IF _n > 0 THEN
    _n          := _n - 1;
    stsVerified := FALSE;
    IF _n = 0 THEN
        _state := E_CamTeach_State.eIdle;
    ELSE
        _state := eTeaching;
    END_IF
END_IF
cmdDeleteLast := TRUE;
END_METHOD

// Spot-edit one existing point (offline, before convert/download). Clears verified.
// Faults on an out-of-range index. Rejected QUIETLY while busy/errored.
METHOD PUBLIC cmdEditPoint : BOOL
VAR_INPUT
    idx     : INT;     // 1..stsNumPoints
    rMaster : LREAL;   // [master unit] new master value
    rSlave  : LREAL;   // [slave unit]  new slave value
END_VAR
cmdEditPoint := FALSE;
IF isBusy() OR stsError THEN
    RETURN;
END_IF

IF idx < 1 OR idx > _n THEN
    setError('Edit point: index out of range');
    RETURN;
END_IF

_points[idx].rMaster := rMaster;
_points[idx].rSlave  := rSlave;
stsVerified  := FALSE;
_state       := eTeaching;
cmdEditPoint := TRUE;
END_METHOD

// Empty the working set (returns toward E_CamTeach_State.eIdle). Clears verified. Rejected QUIETLY while busy/errored.
METHOD PUBLIC cmdClear : BOOL
cmdClear := FALSE;
IF isBusy() OR stsError THEN
    RETURN;
END_IF

_n          := 0;
stsVerified := FALSE;
_state      := E_CamTeach_State.eIdle;
cmdClear    := TRUE;
END_METHOD

// Persist the raw points -> file (async, via fb_CamTeachFile). The directory is cfgFileDir;
// the caller passes just a bare file name. Metadata (slaveName/created/periodic/interp/masterUnit)
// is taken from the cfg backing except 'created', which the HMI stamps (wall clock not in-scan).
// Rejected QUIETLY while busy/errored or with nothing to save.
METHOD PUBLIC cmdSave : BOOL
VAR_INPUT
    fileName : STRING;   // bare file name, e.g. '<pattern>_<slaveName>.csv'
END_VAR
VAR
    sInterp : STRING;
END_VAR
cmdSave := FALSE;
IF isBusy() OR stsError THEN
    RETURN;
END_IF

IF _n < 1 THEN
    setError('Save: nothing to save');
    RETURN;
END_IF

// string form of the interpolation strategy for the CSV '#' header
sInterp := SEL(_interp = E_CamTeach_Interp.eCubicC1, 'linear', 'cubicC1');

IF _file.cmdSave(
        dir        := _fileDir,
        fileName   := fileName,
        numPoints  := _n,
        slaveName  := _slaveName,
        created    := HMI.Config.created,
        periodic   := _periodic,
        interp     := sInterp,
        masterUnit := _masterUnit) THEN
    _fileName    := fileName;
    _returnState := _state;         // resting state to return to once the write completes
    _state       := eSaving;
    cmdSave      := TRUE;
END_IF
END_METHOD

// File -> raw points (async, via fb_CamTeachFile). On completion _n is taken from
// _file.stsNumPointsLoaded and validated (>= 2) in the eLoading branch of the body.
// Loading invalidates any verified table. Rejected QUIETLY while busy/errored.
METHOD PUBLIC cmdLoad : BOOL
VAR_INPUT
    fileName : STRING;   // bare file name to load (directory is cfgFileDir)
END_VAR
cmdLoad := FALSE;
IF isBusy() OR stsError THEN
    RETURN;
END_IF

IF _file.cmdLoad(dir := _fileDir, fileName := fileName) THEN
    _fileName := fileName;
    _state    := eLoading;
    cmdLoad   := TRUE;
END_IF
END_METHOD

// SYNCHRONOUS: post-process the raw points then build the NC motion function _mfPoints[].
// Pure and bounded by MAX_CAM_POINTS (no I/O), so it completes in one scan -> eConverted.
// Post-processing is IN PLACE (design doc "compact the array"): it zeroes the master offset,
// deletes non-monotonic points, and optionally smooths the master column, updating _n. Save
// the raw points BEFORE converting if the untouched values are needed. A (re)convert also
// invalidates any prior download (stsVerified := FALSE). Rejected QUIETLY while busy/errored.
METHOD PUBLIC cmdConvert : BOOL
VAR
    base : LREAL;   // master offset removed in step 1
    i    : INT;     // point loop index
    j    : INT;     // compaction write cursor
    w2   : INT;     // smoothing half-window
    lo   : INT;     // smoothing window low bound
    hi   : INT;     // smoothing window high bound
    k    : INT;     // smoothing inner index
    sum  : LREAL;   // smoothing accumulator
END_VAR
cmdConvert := FALSE;
IF isBusy() OR stsError THEN
    RETURN;
END_IF

IF _n < 2 THEN
    setError('Convert: need at least 2 taught points');
    RETURN;
END_IF

// A (re)convert invalidates any previously downloaded/verified table.
stsVerified := FALSE;

// ── Post-processing 1: zero the master offset (table starts at master = 0) ──
base := _points[1].rMaster;
FOR i := 1 TO _n DO
    _points[i].rMaster := _points[i].rMaster - base;
END_FOR

// ── Post-processing 2: enforce strict-monotonic master (compact the array in place) ──
// Keep point 1; keep each later point only if its master exceeds the last kept point's.
j := 1;
FOR i := 2 TO _n DO
    IF _points[i].rMaster > _points[j].rMaster THEN
        j := j + 1;
        _points[j] := _points[i];
    END_IF
END_FOR
_n := j;
IF _n < 2 THEN
    setError('Convert: too few monotonic points');
    RETURN;
END_IF

// ── Post-processing 3: optional moving-average smoothing of the MASTER column ──
// Odd window (>= 3); the window shrinks at the endpoints. _mfPoints[].MasterPos is used as
// scratch so each average is taken from the ORIGINAL masters (an in-place average would feed
// already-smoothed neighbours into later points). 0/1/2 disable smoothing.
IF _smoothWindow >= 3 THEN
    w2 := (_smoothWindow - 1) / 2;
    FOR i := 1 TO _n DO
        lo := i - w2;  IF lo < 1  THEN lo := 1;  END_IF
        hi := i + w2;  IF hi > _n THEN hi := _n; END_IF
        sum := 0.0;
        FOR k := lo TO hi DO
            sum := sum + _points[k].rMaster;
        END_FOR
        _mfPoints[i].MasterPos := sum / INT_TO_LREAL(hi - lo + 1);   // scratch (overwritten below)
    END_FOR
    FOR i := 1 TO _n DO
        _points[i].rMaster := _mfPoints[i].MasterPos;
    END_FOR
END_IF

// ── Build the NC motion function (C1-smooth cubic from position-only teaching) ──
// Field names and enums checked against TF5050 manual 1.9.2 (section 9.7-9.10), 2026-10-18.
// PointType MUST be set: its default 0 is MOTIONPOINTTYPE_IGNORE, and a table of ignored points is
// rejected (NC 0x4A23 'Motion Function has too few points'). Segments are POLYNOM3_VV (velo <-> velo:
// a cubic through each point's position AND slope) - plain POLYNOM3 is rest <-> rest, i.e. the slave
// would stop at every taught point whatever SlaveVelo says.
FOR i := 1 TO _n DO
    _mfPoints[i].PointIndex        := INT_TO_UDINT(i);       // 1, 2, 3 ... (> 0, consecutive, no gaps)
    _mfPoints[i].PointType         := MOTIONPOINTTYPE_MOTION;
    _mfPoints[i].RelIndexNextPoint := 1;
    _mfPoints[i].MasterPos         := _points[i].rMaster;
    _mfPoints[i].SlavePos          := _points[i].rSlave;
    _mfPoints[i].SlaveVelo         := slaveSlope(i);         // dSlave/dMaster at this point
    _mfPoints[i].SlaveAcc          := 0.0;
    _mfPoints[i].SlaveJerk         := 0.0;
    IF i = _n THEN
        _mfPoints[i].FunctionType      := MOTIONFUNCTYPE_NOTDEF; // last point: no segment after it
        _mfPoints[i].RelIndexNextPoint := 0;                     // ... and no next point (1 -> index _n+1, NC 0x4A13?)
    ELSE
        _mfPoints[i].FunctionType := MOTIONFUNCTYPE_POLYNOM3_VV; // segment to the next point
    END_IF
END_FOR

_state     := eConverted;
cmdConvert := TRUE;
END_METHOD

// Start the async download -> verify state machine (MC_CamTableSelect creates the table, then per-point
// MC_ReadMotionFunctionPoint read-back). On success -> eVerified + stsVerified := TRUE. Requires
// eConverted and a bound cfgTableId. Rejected QUIETLY while busy/errored.
METHOD PUBLIC cmdDownload : BOOL
cmdDownload := FALSE;
IF isBusy() OR stsError THEN
    RETURN;
END_IF

IF _state <> eConverted THEN
    setError('Download: convert first (must be in eConverted)');
    RETURN;
END_IF

IF _tableId = 0 THEN
    setError('Download: no NC cam table id configured');
    RETURN;
END_IF

IF _n < 2 THEN
    setError('Download: nothing to download');
    RETURN;
END_IF

stsVerified := FALSE;               // clears any prior verify until this download re-verifies
_dlStep     := 0;
_state      := eDownloading;
cmdDownload := TRUE;
END_METHOD

// Live single-point slave edit while the table is in use. Updates _points[idx].rSlave, rebuilds
// the affected motion-function points (the edited point's SlavePos + the slopes of it and its
// immediate neighbours), then kicks the async sequence: set the online-change mode (apply at a
// defined master position, NOT immediately) and write the affected points via
// MC_WriteMotionFunctionPoint. The file is re-saved so it stays truthful. A live edit clears
// stsVerified (a full re-convert + re-download is required before coupling is allowed again).
// Rejected QUIETLY while busy/errored, on a bad index, or with no bound table.
METHOD PUBLIC cmdEditOnline : BOOL
VAR_INPUT
    idx    : INT;     // 1..stsNumPoints target point index
    rSlave : LREAL;   // [slave unit] new slave value for the live edit
END_VAR
VAR
    k  : INT;
    lo : INT;
    hi : INT;
END_VAR
cmdEditOnline := FALSE;
IF isBusy() OR stsError THEN
    RETURN;
END_IF

IF _n < 2 THEN
    setError('Online edit: table too small');
    RETURN;
END_IF

IF idx < 1 OR idx > _n THEN
    setError('Online edit: index out of range');
    RETURN;
END_IF

IF _tableId = 0 THEN
    setError('Online edit: no NC cam table id configured');
    RETURN;
END_IF

// 1) update the working point and rebuild the affected motion-function points
//    (only the slave changed; recompute SlavePos of idx and the slopes of idx-1..idx+1).
_onlineIdx := idx;
_points[idx].rSlave := rSlave;

lo := idx - 1;  IF lo < 1  THEN lo := 1;  END_IF
hi := idx + 1;  IF hi > _n THEN hi := _n; END_IF
FOR k := lo TO hi DO
    _mfPoints[k].SlavePos  := _points[k].rSlave;    // VERIFY: MC_MotionFunctionPoint.SlavePos
    _mfPoints[k].SlaveVelo := slaveSlope(k);        // VERIFY: MC_MotionFunctionPoint.SlaveVelo
END_FOR

// 2) + 3) arm the async write sequence: change-mode first, then write points lo..hi.
_onlineWriteIdx := lo;
_onlineHi       := hi;
_onlineStep     := 10;
_onlineSaveReq  := TRUE;

// 4) a live edit invalidates the verified permission; report the updated-but-unverified state.
stsVerified := FALSE;
_state      := eConverted;

cmdEditOnline := TRUE;
END_METHOD

// Clear the FB's own error, reset the file sub-FB, and return to E_CamTeach_State.eIdle. Also aborts any in-flight
// download/verify/online sequence. stsVerified is cleared so a fresh convert + download + verify
// is required after a reset. Called from inpReset, ocmdReset, and directly.
METHOD PUBLIC cmdReset : BOOL
stsError     := FALSE;
stsErrorText := '';
_file.cmdReset();

_state          := E_CamTeach_State.eIdle;
_dlStep         := 0;
_verifyIdx      := 1;
_onlineStep     := 0;
_onlineWriteIdx := 1;
_onlineSaveReq  := FALSE;
stsVerified     := FALSE;
cmdReset        := TRUE;
END_METHOD

// Central-difference slave slope d(slave)/d(master) at point idx, used for the cubic SlaveVelo.
// Interior points use the central difference; the endpoints use one-sided differences. For a
// PERIODIC table the seam (point 1 == point _n phase) wraps so the slope is continuous across
// the period boundary. Assumes masters are strictly monotonic (post-processed); guards dM = 0.
METHOD PRIVATE slaveSlope : LREAL
VAR_INPUT
    idx : INT;     // 1.._n
END_VAR
VAR
    dM     : LREAL;
    dS     : LREAL;
    period : LREAL;
END_VAR
slaveSlope := 0.0;
IF _n < 2 OR idx < 1 OR idx > _n THEN
    RETURN;
END_IF

IF _periodic AND _n >= 3 AND (idx = 1 OR idx = _n) THEN
    // Seam wrap: _points[1] (master 0) and _points[_n] (master = period) are the SAME phase,
    // so idx=1 and idx=_n get the SAME (continuous) slope. period = the zeroed master span.
    period := _points[_n].rMaster - _points[1].rMaster;
    dS     := _points[2].rSlave - _points[_n - 1].rSlave;
    dM     := (_points[2].rMaster + period) - _points[_n - 1].rMaster;
ELSIF idx = 1 THEN
    // one-sided forward difference at the start
    dS := _points[2].rSlave  - _points[1].rSlave;
    dM := _points[2].rMaster - _points[1].rMaster;
ELSIF idx = _n THEN
    // one-sided backward difference at the end
    dS := _points[_n].rSlave  - _points[_n - 1].rSlave;
    dM := _points[_n].rMaster - _points[_n - 1].rMaster;
ELSE
    // interior central difference
    dS := _points[idx + 1].rSlave  - _points[idx - 1].rSlave;
    dM := _points[idx + 1].rMaster - _points[idx - 1].rMaster;
END_IF

IF dM <> 0.0 THEN
    slaveSlope := dS / dM;
END_IF
END_METHOD

// Latch the FB's own error (this FB does NOT extend abs_fb_Device - never setFault, which would
// gate MC_Power on a real axis). Moves to E_CamTeach_State.eError and aborts any in-flight download/verify/online
// sub-steps so the MC blocks de-assert next scan. Cleared only by cmdReset / inpReset.
METHOD PRIVATE setError : BOOL
VAR_INPUT
    text : STRING;
END_VAR
stsError     := TRUE;
stsErrorText := text;
_state       := E_CamTeach_State.eError;
_dlStep      := 0;
_onlineStep  := 0;
setError     := TRUE;
END_METHOD

// TRUE while any async operation is in progress (file save/load, download, verify, or online
// edit). Command methods use this to reject re-entrant requests without disturbing the running op.
METHOD PRIVATE isBusy : BOOL
isBusy := _file.stsBusy
    OR (_state = eSaving) OR (_state = eLoading)
    OR (_state = eDownloading) OR (_state = eVerifying)
    OR (_onlineStep <> 0);
END_METHOD

// Return the full HMI interface struct (the one an HMI binds).
METHOD PUBLIC getHMIdata : ST_CamTeach_HMI_Interface
getHMIdata := HMI;
END_METHOD

METHOD FB_Init : BOOL
VAR_INPUT
    bInitRetains    : BOOL;
    bInCopyCode     : BOOL;
    cfgTableId      : UDINT;              // NC motion-function table id bound to this instance
    cfgSlaveName    : STRING;             // name of the slave this table teaches (file header)
    cfgPeriodic     : BOOL;              // TRUE = periodic table (velocity wraps at the seam)
    cfgInterp       : E_CamTeach_Interp;  // interpolation strategy for cmdConvert
    cfgSmoothWindow : INT;               // moving-average window on master column (0 = off)
    cfgFileDir      : STRING;            // save/load directory ('' = keep default C:\_MachineConfig\CamTables)
    cfgMasterUnit   : STRING;            // CSV header master unit ('' = keep default 'mm')
END_VAR
_tableId   := cfgTableId;
_slaveName := cfgSlaveName;
_periodic  := cfgPeriodic;
_interp    := cfgInterp;
IF cfgSmoothWindow >= 0 THEN _smoothWindow := cfgSmoothWindow; END_IF
IF cfgFileDir    <> '' THEN _fileDir    := cfgFileDir;    END_IF
IF cfgMasterUnit <> '' THEN _masterUnit := cfgMasterUnit; END_IF
END_METHOD

// NC motion-function table id this instance downloads to (pre-created under Motion -> Tables).
PROPERTY PUBLIC cfgTableId : UDINT
GET
cfgTableId := _tableId;
END_GET
SET
_tableId := cfgTableId;
END_SET
END_PROPERTY

// Name of the slave this table teaches; written into the CSV '#' metadata header.
PROPERTY PUBLIC cfgSlaveName : STRING
GET
cfgSlaveName := _slaveName;
END_GET
SET
_slaveName := cfgSlaveName;
END_SET
END_PROPERTY

// TRUE = periodic table: the conversion wraps the central-difference slope at the seam so the
// slave velocity is continuous across the period boundary.
PROPERTY PUBLIC cfgPeriodic : BOOL
GET
cfgPeriodic := _periodic;
END_GET
SET
_periodic := cfgPeriodic;
END_SET
END_PROPERTY

// Interpolation strategy used by cmdConvert (eLinear / eCubicC1). eCubicC1 = POLYNOM3 +
// central-difference slope -> C1-smooth cubic from position-only teaching.
PROPERTY PUBLIC cfgInterp : E_CamTeach_Interp
GET
cfgInterp := _interp;
END_GET
SET
_interp := cfgInterp;
END_SET
END_PROPERTY

// Moving-average window applied to the master column in cmdConvert (odd, 3-5; 0 = off).
// A value < 0 is rejected; 1/2 act as off (the convert only smooths for windows >= 3).
PROPERTY PUBLIC cfgSmoothWindow : INT
GET
cfgSmoothWindow := _smoothWindow;
END_GET
SET
IF cfgSmoothWindow >= 0 THEN _smoothWindow := cfgSmoothWindow; END_IF
END_SET
END_PROPERTY

// Save/load directory (the caller passes only a bare file name). Default C:\_MachineConfig\CamTables.
PROPERTY PUBLIC cfgFileDir : STRING
GET
cfgFileDir := _fileDir;
END_GET
SET
IF cfgFileDir <> '' THEN _fileDir := cfgFileDir; END_IF
END_SET
END_PROPERTY

// Master unit label written into the CSV '#' header (e.g. 'mm' / 'deg'). Default 'mm'.
// Added beyond the design doc's cfg list because the file header needs a machine-specific
// master unit that fb_CamTeachFile.cmdSave requires (see the FB header note / report).
PROPERTY PUBLIC cfgMasterUnit : STRING
GET
cfgMasterUnit := _masterUnit;
END_GET
SET
IF cfgMasterUnit <> '' THEN _masterUnit := cfgMasterUnit; END_IF
END_SET
END_PROPERTY

END_FUNCTION_BLOCK

// ---- POUs/FBs/Camming/fb_CamTeachFile.TcPOU
// fb_CamTeachFile - isolated async CSV persistence for ONE cam-teach table.
//
// Standalone library primitive: does NOT extend abs_fb_Device. It carries its own
// error model (stsError / stsErrorId / stsErrorText) and is driven cyclically by
// fb_CamTeach, which passes its working point array in via VAR_IN_OUT every scan.
//
// The body mirrors the Tc2_System FB_File* async pattern (see fb_WriteDataToFile):
// FB_FileOpen -> FB_FilePuts / FB_FileGets -> FB_FileClose, sequenced by an nState
// CASE machine. Every step is non-blocking (one line per scan pass) and the error
// path (900..) ALWAYS closes the handle before halting.
//
// Operations are started ONLY from cmdSave / cmdLoad, and only when idle (nState = 0),
// so the body never self-triggers. The file is the source of truth; store RAW points.
//
// CSV format (raw values):
//   # slaveName=..  created=..  numPoints=..  periodic=0|1  interp=..  masterUnit=..
//   <master>, <slave>
//   ...
FUNCTION_BLOCK fb_CamTeachFile
VAR_IN_OUT
    // Shared working buffer owned by fb_CamTeach (passed in every scan).
    // Save reads points[1..numPoints]; Load overwrites points[1..stsNumPointsLoaded].
    points : ARRAY[1..MAX_CAM_POINTS] OF ST_CamTeach_Point;
END_VAR
VAR_OUTPUT
    stsBusy            : BOOL;    // an async save/load is in progress
    stsDone            : BOOL;    // last operation finished OK (latched until next op / cmdReset)
    stsError           : BOOL;    // last operation failed (latched until cmdReset)
    stsErrorId         : UDINT;   // Tc2 file-FB error id (nErrId) of the failing step, else 0
    stsErrorText       : STRING;  // human-readable failure description
    stsNumPointsLoaded : INT;     // number of points loaded by the last cmdLoad
END_VAR
VAR
    nState        : INT;          // 0 idle; 10.. save; 110.. load; 900.. error

    // Tc2_System line-oriented file blocks (async; one line per FB_FilePuts/FB_FileGets)
    fbFileOpen    : FB_FileOpen;
    fbFilePuts    : FB_FilePuts;
    fbFileGets    : FB_FileGets;
    fbFileClose   : FB_FileClose;
    hFile         : UINT := 0;    // open file handle (0 = closed)

    // Operation parameters captured by cmdSave / cmdLoad
    _dir          : STRING(255);
    _fileName     : STRING(255);
    _slaveName    : STRING;
    _created      : STRING;
    _interp       : STRING;
    _masterUnit   : STRING;
    _numPoints    : INT;          // points to save (from cmdSave)
    _periodic     : BOOL;

    // Working scratch
    sFullFilePath : STRING(255);  // dir + '\' + fileName
    sLine         : STRING(255);  // line buffer (built for puts / trimmed from gets)
    _i            : INT;          // save row cursor
    _n            : INT;          // load row count
    _hdrNumPoints : INT;          // numPoints parsed from the '#' header (0 = not found)
    rMaster       : LREAL;        // parseRow output scratch
    rSlave        : LREAL;        // parseRow output scratch
END_VAR

CASE nState OF

// ── 0. Idle ─────────────────────────────────────────────────────────────────────
    0:
        stsBusy := FALSE;
        // stsDone / stsError latch until the next command / cmdReset (not cleared here).

// ══ SAVE ═════════════════════════════════════════════════════════════════════════
// ── 10. Build path, open file for writing ────────────────────────────────────────
    10:
        sFullFilePath := _dir;
        IF RIGHT(sFullFilePath, 1) <> '\' THEN
            sFullFilePath := CONCAT(sFullFilePath, '\');   // caller may or may not pass a trailing '\'
        END_IF
        sFullFilePath := CONCAT(sFullFilePath, _fileName);
        fbFileOpen(
            bExecute  := TRUE,
            sNetId    := '',
            sPathName := sFullFilePath,
            nMode     := FOPEN_MODEWRITE OR FOPEN_MODETEXT,
            ePath     := PATH_GENERIC,
            tTimeout  := T#5S);
        nState := 20;

// ── 20. Wait for open ────────────────────────────────────────────────────────────
    20:
        fbFileOpen(bExecute := FALSE);
        IF NOT fbFileOpen.bBusy THEN
            IF fbFileOpen.bError THEN
                stsErrorId   := fbFileOpen.nErrId;
                stsErrorText := 'File open failed (save)';
                nState       := 900;
            ELSE
                hFile  := fbFileOpen.hFile;
                nState := 30;
            END_IF
        END_IF

// ── 30. Write the '#' metadata header line ───────────────────────────────────────
    30:
        sLine := '# slaveName=';
        sLine := CONCAT(sLine, _slaveName);
        sLine := CONCAT(sLine, '  created=');
        sLine := CONCAT(sLine, _created);
        sLine := CONCAT(sLine, '  numPoints=');
        sLine := CONCAT(sLine, INT_TO_STRING(_numPoints));
        sLine := CONCAT(sLine, '  periodic=');
        sLine := CONCAT(sLine, SEL(_periodic, '0', '1'));   // FALSE -> '0', TRUE -> '1'
        sLine := CONCAT(sLine, '  interp=');
        sLine := CONCAT(sLine, _interp);
        sLine := CONCAT(sLine, '  masterUnit=');
        sLine := CONCAT(sLine, _masterUnit);
        sLine := CONCAT(sLine, '$N');
        // VERIFY: FB_FilePuts line-ending behavior is TC-version-dependent. We append LF
        // ('$N') so rows are never concatenated onto one line. If your Tc2_System FB_FilePuts
        // already appends CR/LF, drop this '$N' to avoid blank lines between rows (the loader
        // skips blank lines regardless, so a mismatch degrades cosmetics, not correctness).
        fbFilePuts(bExecute := TRUE, sNetId := '', hFile := hFile, sLine := sLine, tTimeout := T#5S);
        nState := 40;

// ── 40. Wait for header write, arm the row loop ─────────────────────────────────
    40:
        fbFilePuts(bExecute := FALSE);
        IF NOT fbFilePuts.bBusy THEN
            IF fbFilePuts.bError THEN
                stsErrorId   := fbFilePuts.nErrId;
                stsErrorText := 'File write failed (header)';
                nState       := 900;
            ELSE
                _i     := 1;
                nState := 50;
            END_IF
        END_IF

// ── 50. Write one data row (loops 50<->60 until all points written) ──────────────
    50:
        IF _i > _numPoints THEN
            nState := 70;                       // all rows written -> close
        ELSE
            sLine := LREAL_TO_STRING(points[_i].rMaster);
            sLine := CONCAT(sLine, ', ');
            sLine := CONCAT(sLine, LREAL_TO_STRING(points[_i].rSlave));
            sLine := CONCAT(sLine, '$N');       // see VERIFY note in state 30
            fbFilePuts(bExecute := TRUE, sNetId := '', hFile := hFile, sLine := sLine, tTimeout := T#5S);
            nState := 60;
        END_IF

// ── 60. Wait for row write, advance cursor ──────────────────────────────────────
    60:
        fbFilePuts(bExecute := FALSE);
        IF NOT fbFilePuts.bBusy THEN
            IF fbFilePuts.bError THEN
                stsErrorId   := fbFilePuts.nErrId;
                stsErrorText := 'File write failed (row)';
                nState       := 900;
            ELSE
                _i     := _i + 1;
                nState := 50;                   // next row
            END_IF
        END_IF

// ── 70. Close file (save success) ───────────────────────────────────────────────
    70:
        fbFileClose(bExecute := TRUE, sNetId := '', hFile := hFile, tTimeout := T#5S);
        nState := 80;

// ── 80. Wait for close -> Done ──────────────────────────────────────────────────
    80:
        fbFileClose(bExecute := FALSE);
        IF NOT fbFileClose.bBusy THEN
            hFile := 0;
            IF fbFileClose.bError THEN
                stsErrorId   := fbFileClose.nErrId;
                stsErrorText := 'File close failed (save)';
                nState       := 900;
            ELSE
                stsBusy := FALSE;
                stsDone := TRUE;
                nState  := 0;
            END_IF
        END_IF

// ══ LOAD ═════════════════════════════════════════════════════════════════════════
// ── 110. Build path, open file for reading ───────────────────────────────────────
    110:
        sFullFilePath := _dir;
        IF RIGHT(sFullFilePath, 1) <> '\' THEN
            sFullFilePath := CONCAT(sFullFilePath, '\');
        END_IF
        sFullFilePath := CONCAT(sFullFilePath, _fileName);
        fbFileOpen(
            bExecute  := TRUE,
            sNetId    := '',
            sPathName := sFullFilePath,
            nMode     := FOPEN_MODEREAD OR FOPEN_MODETEXT,
            ePath     := PATH_GENERIC,
            tTimeout  := T#5S);
        nState := 120;

// ── 120. Wait for open, init load counters ──────────────────────────────────────
    120:
        fbFileOpen(bExecute := FALSE);
        IF NOT fbFileOpen.bBusy THEN
            IF fbFileOpen.bError THEN
                stsErrorId   := fbFileOpen.nErrId;
                stsErrorText := 'File open failed (load)';
                nState       := 900;
            ELSE
                hFile         := fbFileOpen.hFile;
                _n            := 0;
                _hdrNumPoints := 0;
                nState        := 130;
            END_IF
        END_IF

// ── 130. Read one line ──────────────────────────────────────────────────────────
    130:
        fbFileGets(bExecute := TRUE, sNetId := '', hFile := hFile, tTimeout := T#5S);
        nState := 140;

// ── 140. Classify line: EOF / blank / '#' header / data row (robust) ────────────
    140:
        fbFileGets(bExecute := FALSE);
        IF NOT fbFileGets.bBusy THEN
            IF fbFileGets.bError THEN
                stsErrorId   := fbFileGets.nErrId;
                stsErrorText := 'File read failed (load)';
                nState       := 900;
            ELSIF fbFileGets.bEOF THEN
                nState := 150;                  // end of file -> close
            ELSE
                sLine := fbFileGets.sLine;
                trimWs(sLine);                       // strip CR/LF and surrounding spaces (in place)
                IF sLine = '' THEN
                    nState := 130;              // skip blank lines
                ELSIF LEFT(sLine, 1) = '#' THEN
                    _hdrNumPoints := parseHeaderNumPoints(sLine);   // best-effort count hint
                    nState := 130;              // skip/ignore '#' metadata lines
                ELSE
                    // data row "master, slave"
                    IF parseRow(sLine := sLine, rMaster => rMaster, rSlave => rSlave) THEN
                        IF _n < MAX_CAM_POINTS THEN
                            _n := _n + 1;
                            points[_n].rMaster := rMaster;
                            points[_n].rSlave  := rSlave;
                        END_IF
                    END_IF
                    // stop once the header count is satisfied or the buffer is full;
                    // otherwise keep reading to EOF (robust to a missing/wrong header).
                    IF (_hdrNumPoints > 0 AND _n >= _hdrNumPoints) OR _n >= MAX_CAM_POINTS THEN
                        nState := 150;
                    ELSE
                        nState := 130;
                    END_IF
                END_IF
            END_IF
        END_IF

// ── 150. Close file (load success) ──────────────────────────────────────────────
    150:
        fbFileClose(bExecute := TRUE, sNetId := '', hFile := hFile, tTimeout := T#5S);
        nState := 160;

// ── 160. Wait for close -> Done ─────────────────────────────────────────────────
    160:
        fbFileClose(bExecute := FALSE);
        IF NOT fbFileClose.bBusy THEN
            hFile := 0;
            IF fbFileClose.bError THEN
                stsErrorId   := fbFileClose.nErrId;
                stsErrorText := 'File close failed (load)';
                nState       := 900;
            ELSE
                stsNumPointsLoaded := _n;
                stsBusy := FALSE;
                stsDone := TRUE;
                nState  := 0;
            END_IF
        END_IF

// ══ ERROR PATH (always closes the handle) ════════════════════════════════════════
// ── 900. Enter error, de-assert all file blocks ─────────────────────────────────
    900:
        stsError := TRUE;
        stsBusy  := FALSE;
        fbFileOpen(bExecute := FALSE);
        fbFilePuts(bExecute := FALSE);
        fbFileGets(bExecute := FALSE);
        nState := 910;

// ── 910. Close the handle if still open ─────────────────────────────────────────
    910:
        IF hFile <> 0 THEN
            fbFileClose(bExecute := TRUE, sNetId := '', hFile := hFile, tTimeout := T#5S);
            IF NOT fbFileClose.bBusy THEN
                fbFileClose(bExecute := FALSE);
                hFile  := 0;
                nState := 920;
            END_IF
        ELSE
            nState := 920;
        END_IF

// ── 920. Halt in error - wait for cmdReset ──────────────────────────────────────
    920:
        // latched: stsError stays TRUE until cmdReset() returns the FB to idle.

END_CASE

// Start an async save of points[1..numPoints] to <dir>\<fileName>.
// Guarded: only kicks off when fully idle (nState = 0, not busy, not errored).
// Returns TRUE if accepted, FALSE if rejected (busy/errored - caller should retry
// or cmdReset first). All metadata is copied for the CSV '#' header.
METHOD PUBLIC cmdSave : BOOL
VAR_INPUT
    dir        : STRING(255); // directory (caller's cfgFileDir, e.g. 'C:\_MachineConfig\CamTables')
    fileName   : STRING(255); // bare file name, e.g. '<pattern>_<slaveName>.csv'
    numPoints  : INT;         // number of valid points in points[] to write
    slaveName  : STRING;      // header: name of the slave this table teaches
    created    : STRING;      // header: ISO timestamp supplied by caller/HMI
    periodic   : BOOL;        // header: 0/1 - periodic table flag
    interp     : STRING;      // header: interpolation label, e.g. 'cubicC1' / 'linear'
    masterUnit : STRING;      // header: master unit label, e.g. 'mm' / 'deg'
END_VAR
IF stsBusy OR nState <> 0 THEN
    cmdSave := FALSE;
    RETURN;
END_IF

_dir        := dir;
_fileName   := fileName;
_numPoints  := numPoints;
_slaveName  := slaveName;
_created    := created;
_periodic   := periodic;
_interp     := interp;
_masterUnit := masterUnit;

// clamp the write count to the buffer bound
IF _numPoints < 0 THEN
    _numPoints := 0;
ELSIF _numPoints > MAX_CAM_POINTS THEN
    _numPoints := MAX_CAM_POINTS;
END_IF

stsBusy := TRUE;
stsDone := FALSE;
hFile   := 0;
nState  := 10;      // enter SAVE branch
cmdSave := TRUE;
END_METHOD

// Start an async load of <dir>\<fileName> into points[]. Leading '#' header lines and
// blank lines are skipped; the numPoints header (if present) caps the read, otherwise
// rows are read to EOF. On completion stsNumPointsLoaded holds the count and stsDone
// pulses TRUE. Guarded: only kicks off when idle. Returns TRUE if accepted.
METHOD PUBLIC cmdLoad : BOOL
VAR_INPUT
    dir      : STRING(255);   // directory (caller's cfgFileDir)
    fileName : STRING(255);   // bare file name to load
END_VAR
IF stsBusy OR nState <> 0 THEN
    cmdLoad := FALSE;
    RETURN;
END_IF

_dir      := dir;
_fileName := fileName;

stsNumPointsLoaded := 0;
stsBusy := TRUE;
stsDone := FALSE;
hFile   := 0;
nState  := 110;     // enter LOAD branch
cmdLoad := TRUE;
END_METHOD

// Clear latched done/error state and return to idle. Intended for error recovery.
// If an operation ended in error the handle was already closed by the 910 path, so
// this only clears status. Rejected implicitly if called mid-op via the start guards.
METHOD PUBLIC cmdReset : BOOL
VAR_INPUT
END_VAR
stsBusy      := FALSE;
stsDone      := FALSE;
stsError     := FALSE;
stsErrorId   := 0;
stsErrorText := '';
nState       := 0;
cmdReset     := TRUE;
END_METHOD

// Strip surrounding whitespace and CR/LF from a line. Base Tc2_Standard has no TRIM,
// so this trims manually. Loops are bounded by the string length (<= 255).
// TwinCAT rejects a length-parameterized STRING as a METHOD return type, so this trims the
// string IN PLACE via a VAR_IN_OUT (keeps the full 255 capacity - no truncation to STRING(80)).
METHOD PRIVATE trimWs : BOOL
VAR_IN_OUT
    str : STRING(255);
END_VAR
// trailing CR / LF / space / tab
WHILE LEN(str) > 0 AND (RIGHT(str, 1) = '$R' OR RIGHT(str, 1) = '$L' OR RIGHT(str, 1) = ' ' OR RIGHT(str, 1) = '$T') DO
    str := DELETE(str, 1, LEN(str));   // delete 1 char at the last position
END_WHILE

// leading space / tab
WHILE LEN(str) > 0 AND (LEFT(str, 1) = ' ' OR LEFT(str, 1) = '$T') DO
    str := DELETE(str, 1, 1);          // delete the first char
END_WHILE

trimWs := TRUE;
END_METHOD

// Best-effort parse of "numPoints=<n>" out of a '#' metadata header line.
// Returns 0 if absent - the loader then reads rows until EOF, so 0 is safe.
METHOD PRIVATE parseHeaderNumPoints : INT
VAR_INPUT
    sHeader : STRING(255);
END_VAR
VAR
    nPos   : INT;
    sRest  : STRING(255);
    nSpace : INT;
    sVal   : STRING(255);
END_VAR
parseHeaderNumPoints := 0;

nPos := FIND(sHeader, 'numPoints=');
IF nPos = 0 THEN
    RETURN;
END_IF

// drop chars 1..(nPos+9): the 10-char token 'numPoints=' ends with '=' at nPos+9
sRest := DELETE(sHeader, nPos + 9, 1);
trimWs(sRest);

// value is the first whitespace-delimited token
nSpace := FIND(sRest, ' ');
IF nSpace > 1 THEN
    sVal := LEFT(sRest, nSpace - 1);
ELSE
    sVal := sRest;
END_IF

trimWs(sVal);
parseHeaderNumPoints := STRING_TO_INT(sVal);
END_METHOD

// Parse one "master, slave" CSV data row into two LREALs. Whitespace around each
// field is tolerated. Returns FALSE (and zeroes the outputs) if the line has no comma
// or an empty field, so a malformed row is skipped rather than corrupting the table.
METHOD PRIVATE parseRow : BOOL
VAR_INPUT
    sLine : STRING(255);
END_VAR
VAR_OUTPUT
    rMaster : LREAL;
    rSlave  : LREAL;
END_VAR
VAR
    sWork  : STRING(255);
    nComma : INT;
    sM     : STRING(255);
    sS     : STRING(255);
END_VAR
parseRow := FALSE;
rMaster  := 0;
rSlave   := 0;

sWork := sLine;
trimWs(sWork);
nComma := FIND(sWork, ',');
IF nComma < 2 THEN
    RETURN;                                         // no comma, or nothing before it
END_IF

sM := LEFT(sWork, nComma - 1);                      // text before the comma
sS := MID(sWork, LEN(sWork) - nComma, nComma + 1);  // text after the comma
trimWs(sM);
trimWs(sS);
IF sM = '' OR sS = '' THEN
    RETURN;
END_IF

// VERIFY: string->LREAL conversion name against installed TwinCAT libs.
// STRING_TO_LREAL is provided by Tc2_Standard/Tc2_Utilities on current TC3; if it is
// unavailable, substitute the installed equivalent (e.g. STRING_TO_REAL, lower precision).
rMaster := STRING_TO_LREAL(sM);
rSlave  := STRING_TO_LREAL(sS);
parseRow := TRUE;
END_METHOD

END_FUNCTION_BLOCK

// ---- POUs/FBs/Abstract/abs_fb_Device.TcPOU
FUNCTION_BLOCK ABSTRACT abs_fb_Device
VAR_INPUT
	inpAuto 			: BOOL;
	inpReset 			: BOOL;
	inpInterlockBypass	: BOOL;
	faultMonitor		: POINTER TO fb_FaultMonitor;

END_VAR
VAR_OUTPUT
	stsFaulted 			: BOOL;
	stsFaultDescription : STRING;
END_VAR
VAR
	_deviceName			: STRING;
	_init				: BOOL;	//DO NOT TOGGLE MANUALLY, WILL DUPLICATE ALARM ENTRY
	_initEventClass		: BOOL;
	_enabled			: BOOL;
	_inAuto				: BOOL;
	Interlock			: fb_Interlock;
	_dataInterlock		: st_interlock;
	_deviceFault		: FB_TcAlarm;
	_deviceMsg			: FB_TcMessage;
	_deviceFaultRaised  : BOOL;
	_clear				: BOOL;
	_warnChannels		: ARRAY [1..20] OF STRING;
	_logChannels		: ARRAY [1..20] OF STRING;
	HMIbasedevice		: ST_Device_HMI_Interface;
	_extraFaults		: ARRAY [1..10] OF STRING;
END_VAR

PROPERTY cfgDeviceName : STRING
GET
cfgDeviceName := _deviceName;
END_GET
SET
_deviceName := cfgDeviceName;
END_SET
END_PROPERTY

PROPERTY cfgEnable : BOOL
GET
cfgEnable := _enabled;
END_GET
SET
_enabled := cfgEnable;
END_SET
END_PROPERTY

PROPERTY cfgInitEventClass : Bool
GET
cfgInitEventClass := _initEventClass;
END_GET
SET
_initEventClass := cfgInitEventClass;
END_SET
END_PROPERTY

METHOD cmdReset : BOOL
VAR_INPUT
END_VAR
END_METHOD

METHOD PUBLIC cmdSetInterlock : BOOL
VAR_INPUT
	interlockIndex : INT;
	description : STRING;
	condition: BOOL;
END_VAR
_dataInterlock.conditions[interlockIndex] := condition;
_dataInterlock.descriptions[interlockIndex] := description;
END_METHOD

METHOD PROTECTED DeviceLogic : BOOL
VAR_INPUT
END_VAR
IF NOT _init AND _initEventClass THEN
	_init := TRUE;
	setInit();
END_IF

_inAuto := inpAuto;

Interlock.name 			:= _DeviceName;
Interlock(inpConfig 	:= _dataInterlock, inpGlobalBypass := inpInterlockBypass );

//Fault Handling
IF stsFaulted AND NOT(_deviceFaultRaised) THEN
	_deviceFaultRaised := TRUE;
	_deviceFault.ipArguments.Clear();
	_deviceFault.ipArguments.AddString(_deviceName).AddString(stsFaultDescription);
	_deviceFault.Raise(nTimeStamp :=0);
END_IF

IF NOT(stsFaulted) THEN
	_deviceFaultRaised := FALSE;
	_deviceFault.Clear(0);
END_IF

IF inpReset THEN
	cmdReset();
END_IF

HMIbasedevice.deviceName		  := _devicename;
HMIbasedevice.enabled			  := _enabled;
HMIbasedevice.stsInAuto			  := _inAuto;
HMIbasedevice.interlock 		  := Interlock.getHMIdata();
HMIbasedevice.stsFaulted		  := stsFaulted;
HMIbasedevice.stsFaultDescription := stsFaultDescription;
END_METHOD

//FB_Init is always available implicitly and it is used primarily for initialization.
//The return value is not evaluated. For a specific influence, you can also declare the
//methods explicitly and provide additional code there with the standard initialization
//code. You can evaluate the return value.
METHOD FB_Init: BOOL
VAR_INPUT
    bInitRetains: BOOL; // TRUE: the retain variables are initialized (reset warm / reset cold)
    bInCopyCode: BOOL;  // TRUE: the instance will be copied to the copy code afterward (online change)   
	cfgDeviceName 		: STRING;
	cfgEnable			: BOOL;
	cfgInitEventClass	: BOOL;
END_VAR
THIS^.cfgDeviceName 		:= 		cfgDeviceName; 
THIS^.cfgEnable				:=		cfgEnable;
THIS^.cfgInitEventClass		:= 		cfgInitEventClass;
END_METHOD

METHOD INTERNAL sendLog : BOOL
VAR_INPUT
	message : STRING;
	channel : USINT;
END_VAR
IF message <> _logChannels[channel] THEN
	_logchannels[channel] := message;
	_deviceMsg.CreateEx(TC_Events.absDevice.Logger,0);
	_deviceMsg.ipArguments.AddString(_deviceName).AddString(message);
	_deviceMsg.Send(0);
END_IF
END_METHOD

METHOD INTERNAL sendWarning : BOOL
VAR_INPUT
	message : STRING;
	channel : USINT;
END_VAR
IF message <> _warnChannels[channel] THEN
	_warnChannels[channel] := message;
	_deviceMsg.CreateEx(TC_Events.absDevice.Warning,0);
	_deviceMsg.ipArguments.AddString(_deviceName).AddString(message);
	_deviceMsg.Send(0);	
END_IF
END_METHOD

METHOD INTERNAL setFault : BOOL
VAR_INPUT
	faultState			: BOOL;
	faultDescription	: STRING;
END_VAR
VAR
	i            : DINT;
	alreadyAdded : BOOL;	// per call: was this description already reported as an additional fault?
END_VAR
// alreadyAdded is LOCAL on purpose. It was an FB member that was only cleared when the fault
// was reset, so after one repeated additional fault every later, DIFFERENT one was dropped.
IF faultState THEN
	//if already faulted, send out additional faults as warnings
	IF stsFaulted AND NOT(faultDescription = stsFaultDescription) THEN
		//Check if already added
		FOR i:= 1 TO UPPER_BOUND(_extraFaults,1) DO
			IF faultDescription = _extraFaults[i] THEN
				alreadyAdded := TRUE;
				EXIT;
			END_IF
		END_FOR
		IF NOT alreadyAdded AND (_extraFaults[10] = '') THEN
			sendWarning(CONCAT('Additional Fault - ', faultDescription),20);
			FOR i:= 1 TO UPPER_BOUND(_extraFaults,1) DO
				IF _extraFaults[i] = '' THEN
					_extraFaults[i] := faultDescription;
					EXIT;
				END_IF
			END_FOR
		END_IF
	ELSE
		stsFaulted := TRUE;
		stsFaultDescription := faultDescription;
	END_IF

ELSE
	stsFaulted := FALSE;
	stsFaultDescription := '';
	MEMSET(destAddr := ADR(_extraFaults), fillByte := 0, n:= SIZEOF(_extraFaults));
END_IF
END_METHOD

METHOD INTERNAL setInit : BOOL
VAR_INPUT
END_VAR
IF faultMonitor <> 0 THEN
	faultMonitor^.addDeviceFault(faultStatus := ADR(stsFaulted), faultDescription := ADR(stsFaultDescription), deviceName := ADR(_deviceName));
END_IF
_deviceFault.CreateEx(stEventEntry:=TC_Events.absDevice.Faulted, bWithConfirmation := FALSE, ipSourceInfo := 0);
_deviceMsg.CreateEx(stEventEntry:=TC_events.absDevice.Warning,ipSourceInfo:=0);
_deviceMsg.CreateEx(stEventEntry:=TC_events.absDevice.Logger,ipSourceInfo:=0);
END_METHOD

END_FUNCTION_BLOCK

// ---- POUs/FBs/fb_FaultMonitor.TcPOU
(*
    fb_FaultMonitor — machine-wide list of the devices that are faulted right now.

    Devices register once (abs_fb_Device / abs_fb_stateDevice call addDeviceFault from setInit with
    pointers to their own stsFaulted / stsFaultDescription / device name). Every scan the monitor
    REBUILDS stsFoundFaultDevice / stsFoundFaultDescription from those pointers, so the two lists
    always line up index for index, a cleared fault disappears the scan it clears, and a fault whose
    text changes shows the current text. (It used to add and remove entries by matching the
    description string, which failed once a device blanked its description on reset: the stale
    text stayed in the list for good.)
*)
FUNCTION_BLOCK fb_FaultMonitor
VAR_INPUT
END_VAR

VAR_OUTPUT
    stsFaultActive           : BOOL;
    stsFaultCount            : UINT;                    // number of entries in the two lists below
    stsFoundFaultDevice      : ARRAY[1..150] OF STRING;
    stsFoundFaultDescription : ARRAY[1..150] OF STRING;
END_VAR

VAR
    _deviceFaults            : ARRAY[1..150] OF POINTER TO BOOL;
    _deviceFaultDescriptions : ARRAY[1..150] OF POINTER TO STRING;
    _deviceNames             : ARRAY[1..150] OF POINTER TO STRING;
    _lastCount               : UINT;
END_VAR

scanFaults();

METHOD addDeviceFault : BOOL
VAR_INPUT
    faultStatus         : POINTER TO BOOL;
    faultDescription    : POINTER TO STRING;
    deviceName          : POINTER TO STRING;
END_VAR
VAR
    deviceFaultIndex    : UINT;
END_VAR
addDeviceFault := FALSE;
IF faultStatus = 0 THEN
    RETURN;
END_IF

deviceFaultIndex := getDeviceFaultArrayIndex(faultStatus);
IF deviceFaultIndex <> 0 THEN
    _deviceFaults[deviceFaultIndex]            := faultStatus;
    _deviceFaultDescriptions[deviceFaultIndex] := faultDescription;
    _deviceNames[deviceFaultIndex]             := deviceName;
    addDeviceFault := TRUE;
END_IF
END_METHOD

// Slot for a registration: the slot this device already holds (so registering twice, e.g.
// after an online change re-runs setInit, does not take a second slot), else the first free
// one. 0 = table full.
METHOD PRIVATE getDeviceFaultArrayIndex : UINT
VAR_INPUT
    faultStatus : POINTER TO BOOL;
END_VAR
VAR
    i           : UINT;
END_VAR
getDeviceFaultArrayIndex := 0;
FOR i := 1 TO 150 DO
    IF _deviceFaults[i] = faultStatus THEN
        getDeviceFaultArrayIndex := i;
        RETURN;
    END_IF
END_FOR
FOR i := 1 TO 150 DO
    IF _deviceFaults[i] = 0 THEN
        getDeviceFaultArrayIndex := i;
        RETURN;
    END_IF
END_FOR
END_METHOD

METHOD PRIVATE scanFaults : BOOL
VAR
    i   : UINT;
    n   : UINT;
END_VAR
n := 0;
FOR i := 1 TO 150 DO
    IF _deviceFaults[i] <> 0 THEN
        IF _deviceFaults[i]^ THEN
            n := n + 1;
            IF _deviceNames[i] <> 0 THEN
                stsFoundFaultDevice[n] := _deviceNames[i]^;
            ELSE
                stsFoundFaultDevice[n] := '';
            END_IF
            IF _deviceFaultDescriptions[i] <> 0 THEN
                stsFoundFaultDescription[n] := _deviceFaultDescriptions[i]^;
            ELSE
                stsFoundFaultDescription[n] := '';
            END_IF
        END_IF
    END_IF
END_FOR

// Blank only the tail the previous scan used, not all 150 entries every scan.
FOR i := n + 1 TO _lastCount DO
    stsFoundFaultDevice[i]      := '';
    stsFoundFaultDescription[i] := '';
END_FOR
_lastCount := n;

stsFaultCount  := n;
stsFaultActive := (n > 0);
END_METHOD

END_FUNCTION_BLOCK

// ---- POUs/FBs/fb_Interlock.TcPOU
FUNCTION_BLOCK fb_Interlock
VAR_INPUT
	inpConfig 		: ST_Interlock;
	inpGlobalBypass	: BOOL;
END_VAR

VAR
	i	: INT;
	HMI : ST_Interlock_HMI_Interface;
END_VAR

VAR_OUTPUT
	outInterlockOK	: BOOL;
	stsFirstOut		: STRING;
END_VAR


outInterlockOK := TRUE;
stsFirstOut := '';
IF NOT(inpGlobalBypass) THEN
	FOR i:= 1 TO 10 DO
		IF NOT inpConfig.conditions[i] THEN
			outInterlockOK := FALSE;
			// FIRST-out, not last: only take the text while it is still empty. This assigned on
			// EVERY failing iteration until 2026-07-26, so despite the name it reported the LAST
			// failing condition. An interlock trips the instant one condition drops, and the point of
			// a first-out readout is to name the condition that CAUSED the trip - slot order is
			// authored upstream-first, so slot 1 is the root cause and slot 10 is usually a
			// consequence of it. Reporting the last one pointed the operator at the symptom.
			IF stsFirstOut = '' THEN
				stsFirstOut := inpConfig.descriptions[i];
			END_IF
		END_IF
	END_FOR
END_IF

HMI.stsInterlockOK := outInterlockOK;
HMI.stsConditions := inpConfig.conditions;
HMI.stsInterlockDescriptions := inpConfig.descriptions;

METHOD PUBLIC getHMIdata : ST_Interlock_HMI_Interface
VAR_INPUT
END_VAR
getHMIdata := HMI;
END_METHOD

PROPERTY PUBLIC name : string
GET
name := HMI.stsInterlockName;
END_GET
SET
hmi.stsInterlockName := name;
END_SET
END_PROPERTY

END_FUNCTION_BLOCK

// ---- POUs/FBs/Abstract/abs_fb_MachineFlow.TcPOU
(*  abs_fb_MachineFlow - parallel machine-sequence composer (SFC-style token engine)
    on top of abs_fb_stateDevice.

    A derived FB declares its sequence as DATA in defineFlow() - addStep() for the
    steps, flow()/flowSplit2..3()/flowJoin2..3() (or addTransition() + arcFrom()/
    arcTo() for other shapes) for the relationships - and writes the step BODIES in
    stepActions(), a CASE over the step ids. The engine holds a token per active
    step: a transition fires when ALL its source steps are active AND done AND its
    permissive is TRUE; firing consumes the source tokens and activates all targets.
    Parallel branches, joins, choices (two transitions from one step with opposing
    permissives) and loops are therefore plain data - no flags, no duplicated states.

    Lifecycle (run/abort/retry/reset, interlocks, alarms, HMI commands) is inherited
    unchanged from abs_fb_stateDevice; the base state variable receives the
    transition-firing counter, so the base step timer measures time since the last
    firing (a stall watchdog). Per-step elapsed/timeout clocks run in the engine
    (parallel-safe); a step timeout faults with retry allowed - retry resumes with
    the timed-out step's clock cleared and all tokens in place.

    Usage:
        FUNCTION_BLOCK fb_SEQ_Wash EXTENDS abs_fb_MachineFlow
        Body (first line):       flowLogic();
        STEP IDS ARE `VAR CONSTANT`, NOT VAR. stepActions() dispatches on them with
        CASE, and IEC 61131-3 requires CASE labels to be CONSTANT - a runtime VAR
        holding addStep()'s return value cannot be a label and will not compile. So
        declare them as constants with explicit literal values, `c`-prefixed per
        CONVENTIONS §2 (never a type prefix - `cStepFill`, never `sFill`):

            VAR CONSTANT
                cStepFill : INT := 1;   // ids are assigned in addStep() CALL ORDER
                cStepHeat : INT := 2;
                cStepStir : INT := 3;
            END_VAR

        The constants and the addStep() order must agree, and nothing enforces it -
        inserting a step in the middle silently shifts every later id. addStep()
        returns the id it actually assigned, so guard it:

        Override defineFlow():   IF addStep('Fill tank', T#30S) <> cStepFill THEN
                                     setCfgError('flow: step id drift'); END_IF
                                 ...
                                 setInitialStep(cStepFill);
                                 flowSplit2(cStepFill, cStepHeat, cStepStir);
        Override stepActions():  CASE inpStepId OF cStepFill: ... stepDone(cStepFill); ...

        Transition ids are NOT dispatched on, so they may be plain VAR (`_transLoop`)
        holding what flow()/addTransition() returned - setPermissive() takes a value.
        A step completes via stepDone(id); a DONE step with no outgoing transition
        completes the sequence (setStateLogicDone). Override actionsAbort() for a
        controlled abort ramp (the default clears the tokens and finishes at once).

    Determinism: transitions are evaluated in ascending id order each scan; firing
    consumes tokens, so two transitions competing for one token resolve to the lower
    id. A newly activated step always executes at least one scan before any outgoing
    transition can fire.

    SELF-CONTAINED (CONVENTIONS §5): this FB references no GVL and holds no pointer
    to anything it does not own. A transition's gate is ONE BOOL - where the gate is
    really an fb_Permissive, the machine ANDs stsPermissiveOK in at the setPermissive()
    call, the same way it reports a step with stepDone(). The engine knows only tokens
    and booleans, which is all a token engine should know.

    Capacities are LITERALS, repeated in the array bounds and in every loop that walks
    them - keep those edits together:
      * 64 steps / 64 transitions. 64 is not arbitrary and is the one number NOT free
        to change: the HMI publishes the active/done/visited/fired/permissive masks as
        2 x UDINT (lo = 1..32, hi = 33..64), so raising it breaks that contract and the
        lhmi renderer with it. Widening means new mask members, not a bigger bound.
      * 4 sources / 4 targets per transition (ST_MachineFlow_Transition) - the widest
        AND-split or AND-join a transition can express.
      * 4095-byte stsFlowDef, the exported definition JSON. Truncation is reported, not
        silent (see actionsRun); step and transition NAMES are what consume it.

    HMI: HMIflow (ST_MachineFlow_HMI_Status) carries the token + permissive masks,
    the firing counter and the STATIC definition JSON including each transition's
    condition text (read once, on demand - ADS only, not for cyclic transport); the
    inherited HMIstateLogic carries state/commands. While the sequence runs,
    stsStepDescription is ENGINE-OWNED: the joined active-step names. Name every
    permissive-gated transition - the name is the operator's answer to 'why is this
    step stuck'. Step/transition names must not contain double quotes (def JSON).
*)
FUNCTION_BLOCK ABSTRACT abs_fb_MachineFlow EXTENDS abs_fb_stateDevice
VAR_OUTPUT
    stsActiveNames  : STRING(255);   // ' + '-joined names of the active steps
END_VAR
VAR
    HMIflow         : ST_MachineFlow_HMI_Status;
    _steps          : ARRAY[1..64] OF ST_MachineFlow_Step;
    _trans          : ARRAY[1..64] OF ST_MachineFlow_Transition;
    _stepTimers     : ARRAY[1..64] OF TON;
    _initialSteps   : ARRAY[1..64] OF BOOL;
    _stepCount      : INT;
    _transCount     : INT;
    _initialCount   : INT;
    _defined        : BOOL;
    _fireCount      : INT;    // the base state variable: transition firings this run
    _lastFired      : INT;
    _timeoutStep    : INT;    // step that raised the running step-timeout fault
    _wasRunning     : BOOL;
    _wasFaulted     : BOOL;
    _defLen         : INT;
    _defOverflow    : BOOL;
    _faultedStep    : INT;   // step that raised (or timed out into) the active fault; 0 = none
    _cfgError       : BOOL;
    _cfgErrorText   : STRING(255);
END_VAR

// Default abort: drop all tokens and finish immediately. Override for a
// controlled ramp-down (make devices safe, then call setStateDoneAborting()).
METHOD PROTECTED actionsAbort : BOOL
VAR_INPUT
END_VAR
clearTokens();
setStateDoneAborting();
actionsAbort := TRUE;
END_METHOD

METHOD PROTECTED actionsReset : BOOL
VAR_INPUT
END_VAR
VAR
    t : INT;
END_VAR
clearTokens();
FOR t := 1 TO _transCount DO
    _trans[t].permissive := TRUE;
    _trans[t].fired := FALSE;
END_FOR
_fireCount := 0;
_lastFired := 0;
_timeoutStep := 0;
_faultedStep := 0;
actionsReset := TRUE;
END_METHOD

// The engine scan: per-step clocks/timeouts -> step bodies (once per active
// step) -> transition firing -> done detection. Runs every cycle while Running.
METHOD PROTECTED actionsRun : BOOL
VAR_INPUT
END_VAR
IF _cfgError THEN
    setStateLogicFault(_cfgErrorText, FALSE, 0);
    RETURN;
END_IF
IF _defOverflow THEN
    _defOverflow := FALSE;
    sendWarning('MachineFlow: definition JSON truncated - shorten step/transition names or widen stsFlowDef (4095)');
END_IF

runStepTimers();
IF stsFaulted THEN
    RETURN;   // a step timeout faulted this scan
END_IF
dispatchSteps();
fireTransitions();
checkFlowDone();
actionsRun := TRUE;
END_METHOD

// Declare a step (call from defineFlow()). Returns the step id used by
// stepActions()/stepDone()/the transitions; 0 on capacity error.
// inpDescription = WHAT the step does, shown in the HMI's step popup.
METHOD PROTECTED addStep : INT
VAR_INPUT
    inpName        : STRING(63);
    inpTimeout     : TIME := T#0S;   // T#0S = no timeout; runtime override: setStepTimeout()
    inpDescription : STRING(125) := '';
END_VAR
IF _stepCount >= 64 THEN
    setCfgError('MachineFlow: addStep() capacity exceeded');
    addStep := 0;
    RETURN;
END_IF
_stepCount := _stepCount + 1;
_steps[_stepCount].name := inpName;
_steps[_stepCount].description := inpDescription;
_steps[_stepCount].timeout := inpTimeout;
addStep := _stepCount;
END_METHOD

// Allocate an empty transition (call from defineFlow()); attach steps with
// arcFrom()/arcTo(). The flow*() helpers cover the common shapes.
// inpName is the CONDITION text the HMI shows on the transition bar
// (e.g. 'cycles < 3') - name every permissive so a held gate explains itself.
METHOD PROTECTED addTransition : INT
VAR_INPUT
    inpName : STRING(63) := '';
END_VAR
IF _transCount >= 64 THEN
    setCfgError('MachineFlow: addTransition() capacity exceeded');
    addTransition := 0;
    RETURN;
END_IF
_transCount := _transCount + 1;
_trans[_transCount].name := inpName;
addTransition := _transCount;
END_METHOD

METHOD PRIVATE appendDef : BOOL
VAR_INPUT
    inpText : STRING(255);
END_VAR
VAR
    txtLen : INT;
    k      : INT;
    pSrc   : POINTER TO BYTE;
    pDst   : POINTER TO BYTE;
END_VAR
txtLen := LEN(inpText);
IF txtLen = 0 THEN
    appendDef := TRUE;
    RETURN;
END_IF
IF _defLen + txtLen >= 4095 THEN
    _defOverflow := TRUE;
    RETURN;
END_IF
pSrc := ADR(inpText);
pDst := ADR(HMIflow.stsFlowDef);
pDst := pDst + _defLen;
FOR k := 0 TO txtLen - 1 DO
    pDst[k] := pSrc[k];
END_FOR
_defLen := _defLen + txtLen;
appendDef := TRUE;
END_METHOD

// Add a SOURCE step to a transition (all sources must be done for it to fire).
METHOD PROTECTED arcFrom : BOOL
VAR_INPUT
    inpTrans  : INT;
    inpStepId : INT;
END_VAR
VAR
    a : INT;
END_VAR
IF inpTrans < 1 OR inpTrans > _transCount OR inpStepId < 1 OR inpStepId > 64 THEN
    setCfgError('MachineFlow: arcFrom() bad transition/step id');
    RETURN;
END_IF
FOR a := 1 TO 4 DO
    IF _trans[inpTrans].sources[a] = 0 THEN
        _trans[inpTrans].sources[a] := inpStepId;
        arcFrom := TRUE;
        RETURN;
    END_IF
END_FOR
setCfgError('MachineFlow: arcFrom() arc capacity exceeded');
END_METHOD

// Add a TARGET step to a transition (all targets activate when it fires).
METHOD PROTECTED arcTo : BOOL
VAR_INPUT
    inpTrans  : INT;
    inpStepId : INT;
END_VAR
VAR
    a : INT;
END_VAR
IF inpTrans < 1 OR inpTrans > _transCount OR inpStepId < 1 OR inpStepId > 64 THEN
    setCfgError('MachineFlow: arcTo() bad transition/step id');
    RETURN;
END_IF
FOR a := 1 TO 4 DO
    IF _trans[inpTrans].targets[a] = 0 THEN
        _trans[inpTrans].targets[a] := inpStepId;
        arcTo := TRUE;
        RETURN;
    END_IF
END_FOR
setCfgError('MachineFlow: arcTo() arc capacity exceeded');
END_METHOD

METHOD PRIVATE buildDefJson : BOOL
VAR_INPUT
END_VAR
VAR
    i, t, a, sid : INT;
    firstArc   : BOOL;
    pEnd       : POINTER TO BYTE;
END_VAR
_defLen := 0;
_defOverflow := FALSE;
appendDef('{"v":1,"steps":[');
FOR i := 1 TO _stepCount DO
    IF i > 1 THEN
        appendDef(',');
    END_IF
    appendDef('{"i":');
    appendDef(INT_TO_STRING(i));
    appendDef(',"n":"');
    appendDef(_steps[i].name);
    appendDef('"');
    IF _steps[i].description <> '' THEN
        appendDef(',"d":"');
        appendDef(_steps[i].description);
        appendDef('"');
    END_IF
    // Step TIMEOUT, in ms, and only when one is configured. Static config, so it belongs in the def
    // (read once) rather than in a cyclic member: 64 timeouts polled every scan would cost real
    // bandwidth for numbers that never change. Omitted when T#0S so an untimed step costs 0 bytes of
    // the 4095 - most steps have no timeout.
    IF _steps[i].timeout > T#0S THEN
        appendDef(',"to":');
        appendDef(UDINT_TO_STRING(TIME_TO_UDINT(_steps[i].timeout)));
    END_IF
    IF _initialSteps[i] THEN
        appendDef(',"init":1');
    END_IF
    appendDef('}');
END_FOR
appendDef('],"trans":[');
FOR t := 1 TO _transCount DO
    IF t > 1 THEN
        appendDef(',');
    END_IF
    appendDef('{"id":');
    appendDef(INT_TO_STRING(t));
    IF _trans[t].name <> '' THEN
        appendDef(',"n":"');
        appendDef(_trans[t].name);
        appendDef('"');
    END_IF
    appendDef(',"s":[');
    firstArc := TRUE;
    FOR a := 1 TO 4 DO
        sid := _trans[t].sources[a];
        IF sid > 0 THEN
            IF NOT firstArc THEN
                appendDef(',');
            END_IF
            appendDef(INT_TO_STRING(sid));
            firstArc := FALSE;
        END_IF
    END_FOR
    appendDef('],"t":[');
    firstArc := TRUE;
    FOR a := 1 TO 4 DO
        sid := _trans[t].targets[a];
        IF sid > 0 THEN
            IF NOT firstArc THEN
                appendDef(',');
            END_IF
            appendDef(INT_TO_STRING(sid));
            firstArc := FALSE;
        END_IF
    END_FOR
    appendDef(']}');
END_FOR
appendDef(']}');
pEnd := ADR(HMIflow.stsFlowDef);
pEnd := pEnd + _defLen;
pEnd^ := 0;
buildDefJson := TRUE;
END_METHOD

METHOD PRIVATE checkFlowDone : BOOL
VAR_INPUT
END_VAR
VAR
    i               : INT;
    anyActive       : BOOL;
    allTerminalDone : BOOL;
END_VAR
allTerminalDone := TRUE;
FOR i := 1 TO _stepCount DO
    IF _steps[i].active THEN
        anyActive := TRUE;
        IF NOT _steps[i].done OR _steps[i].hasOutgoing THEN
            allTerminalDone := FALSE;
        END_IF
    END_IF
END_FOR
IF NOT anyActive THEN
    setStateLogicFault('MachineFlow: no active steps while running (check the flow definition)', FALSE, 0);
ELSIF allTerminalDone THEN
    setStateLogicDone();
END_IF
checkFlowDone := TRUE;
END_METHOD

// Drop every token (and this run's history). PROTECTED because overriding actionsAbort() for a
// controlled ramp-down is a documented extension point, and the default it replaces ends with
// clearTokens() + setStateDoneAborting() - a subclass could not reproduce that while this was
// PRIVATE. Safe to expose: clearing mid-RUN is caught on the next scan by checkFlowDone, which
// faults with 'no active steps while running' rather than hanging silently, and during an abort
// actionsRun() is not running so the legitimate use never trips it.
METHOD PROTECTED clearTokens : BOOL
VAR_INPUT
END_VAR
VAR
    i : INT;
END_VAR
FOR i := 1 TO 64 DO
    _steps[i].active := FALSE;
    _steps[i].done := FALSE;
    _steps[i].visited := FALSE;
    _steps[i].entered := FALSE;
    _steps[i].kickTimer := TRUE;
END_FOR
clearTokens := TRUE;
END_METHOD

// Override: declare the sequence graph - RELATIONSHIPS only, no step logic.
// addStep() the steps, then connect them with flow()/flowSplit2..3()/
// flowJoin2..3() (or addTransition() + arcFrom()/arcTo() for other shapes).
// Called once, before the first scan. Default initial step: the first declared
// one (override with setInitialStep(); call it more than once for parallel starts).
METHOD PROTECTED defineFlow : BOOL
VAR_INPUT
END_VAR
END_METHOD

METHOD PRIVATE dispatchSteps : BOOL
VAR_INPUT
END_VAR
VAR
    i         : INT;
    firstScan : BOOL;
END_VAR
FOR i := 1 TO _stepCount DO
    IF _steps[i].active THEN
        firstScan := NOT _steps[i].entered;
        _steps[i].entered := TRUE;
        stepActions(inpStepId := i, inpFirstScan := firstScan);
        // ATTRIBUTE A STEP-RAISED FAULT TO ITS STEP. A step body may check a condition and call
        // setFault() on the inherited state device: that faults the parent state machine, but the
        // fault also belongs to THIS step, and the HMI needs to know which one so the flow chart can
        // colour it red. Checked right after the body runs, and only claimed if nothing else has -
        // a step timeout (runStepTimers) already sets _faultedStep, and the first claim wins so a
        // later step in the same scan cannot steal the attribution.
        IF stsFaulted AND _faultedStep = 0 THEN
            _faultedStep := i;
        END_IF
    END_IF
END_FOR
dispatchSteps := TRUE;
END_METHOD

METHOD PRIVATE finalizeFlow : BOOL
VAR_INPUT
END_VAR
VAR
    t, a, sid : INT;
END_VAR
// default initial step: the first declared one
IF _initialCount = 0 AND _stepCount > 0 THEN
    _initialSteps[1] := TRUE;
    _initialCount := 1;
END_IF
// derive hasOutgoing + validate every arc against the declared steps
FOR t := 1 TO _transCount DO
    FOR a := 1 TO 4 DO
        sid := _trans[t].sources[a];
        IF sid > 0 THEN
            IF sid > _stepCount THEN
                setCfgError('MachineFlow: a transition source references an unknown step');
            ELSE
                _steps[sid].hasOutgoing := TRUE;
            END_IF
        END_IF
        sid := _trans[t].targets[a];
        IF sid > _stepCount THEN
            setCfgError('MachineFlow: a transition target references an unknown step');
        END_IF
    END_FOR
END_FOR
buildDefJson();
HMIflow.stsStepCount := _stepCount;
HMIflow.stsTransCount := _transCount;
finalizeFlow := TRUE;
END_METHOD

METHOD PRIVATE fireTransitions : BOOL
VAR_INPUT
END_VAR
VAR
    t, a, sid   : INT;
    enabled   : BOOL;
    hasSource : BOOL;
END_VAR
FOR t := 1 TO _transCount DO
    // A transition gate is ONE BOOL, and the engine knows nothing else about it. Where the gate is a
    // full fb_Permissive, the machine ANDs it in at the call site - setPermissive(t,
    // PermUnload.stsPermissiveOK) - exactly as it reports a step with stepDone(id). See the header:
    // this engine holds no reference to anything outside itself.
    enabled := _trans[t].permissive;
    hasSource := FALSE;
    FOR a := 1 TO 4 DO
        sid := _trans[t].sources[a];
        IF sid > 0 THEN
            hasSource := TRUE;
            IF NOT (_steps[sid].active AND _steps[sid].done) THEN
                enabled := FALSE;
            END_IF
        END_IF
    END_FOR
    IF enabled AND hasSource THEN
        // consume every source token first (a self-loop re-places below)
        FOR a := 1 TO 4 DO
            sid := _trans[t].sources[a];
            IF sid > 0 THEN
                _steps[sid].active := FALSE;
                _steps[sid].done := FALSE;
                // Consuming a token IS the moment a step completed. Recorded because the token is
                // gone next scan, leaving nothing to distinguish "finished" from "never ran" - which
                // the flow chart colours differently.
                _steps[sid].visited := TRUE;
            END_IF
        END_FOR
        FOR a := 1 TO 4 DO
            sid := _trans[t].targets[a];
            IF sid > 0 THEN
                placeToken(sid);
            END_IF
        END_FOR
        _lastFired := t;
        _trans[t].fired := TRUE;   // this run; _lastFired only ever holds the newest
        _fireCount := _fireCount + 1;
    END_IF
END_FOR
fireTransitions := TRUE;
END_METHOD

// Simple arrow: source done -> target activates. Returns the transition id
// (keep it to attach a runtime permissive via setPermissive(), e.g. for loop-back edges).
// inpName = the condition text shown on the HMI bar.
METHOD PROTECTED flow : INT
VAR_INPUT
    inpFrom : INT;
    inpTo   : INT;
    inpName : STRING(63) := '';
END_VAR
flow := addTransition(inpName := inpName);
IF flow = 0 THEN
    RETURN;
END_IF
arcFrom(inpTrans := flow, inpStepId := inpFrom);
arcTo(inpTrans := flow, inpStepId := inpTo);
END_METHOD

// AND-convergence: fires when BOTH sources are done; activates the target.
METHOD PROTECTED flowJoin2 : INT
VAR_INPUT
    inpFrom1 : INT;
    inpFrom2 : INT;
    inpTo    : INT;
    inpName  : STRING(63) := '';
END_VAR
flowJoin2 := addTransition(inpName := inpName);
IF flowJoin2 = 0 THEN
    RETURN;
END_IF
arcFrom(inpTrans := flowJoin2, inpStepId := inpFrom1);
arcFrom(inpTrans := flowJoin2, inpStepId := inpFrom2);
arcTo(inpTrans := flowJoin2, inpStepId := inpTo);
END_METHOD

// AND-convergence: fires when ALL THREE sources are done; activates the target.
METHOD PROTECTED flowJoin3 : INT
VAR_INPUT
    inpFrom1 : INT;
    inpFrom2 : INT;
    inpFrom3 : INT;
    inpTo    : INT;
    inpName  : STRING(63) := '';
END_VAR
flowJoin3 := addTransition(inpName := inpName);
IF flowJoin3 = 0 THEN
    RETURN;
END_IF
arcFrom(inpTrans := flowJoin3, inpStepId := inpFrom1);
arcFrom(inpTrans := flowJoin3, inpStepId := inpFrom2);
arcFrom(inpTrans := flowJoin3, inpStepId := inpFrom3);
arcTo(inpTrans := flowJoin3, inpStepId := inpTo);
END_METHOD

// Call as the FIRST line of the derived FB's body (like DeviceLogic() in
// abs_fb_Device). Builds the graph once, handles run/resume edges, then runs
// the inherited state logic (which calls actionsRun = the engine scan).
METHOD PROTECTED flowLogic : BOOL
VAR_INPUT
END_VAR
IF NOT _defined THEN
    _defined := TRUE;
    defineFlow();
    finalizeFlow();
END_IF

// Run/resume edge: a fresh run seeds the initial tokens; a retry-resume keeps
// the tokens in place and only restarts the timed-out step's clock.
IF stsRunning AND NOT _wasRunning THEN
    IF _wasFaulted THEN
        IF _timeoutStep > 0 THEN
            _steps[_timeoutStep].kickTimer := TRUE;
            _timeoutStep := 0;
_faultedStep := 0;
        END_IF
    ELSE
        seedTokens();
    END_IF
END_IF
_wasRunning := stsRunning;
_wasFaulted := stsFaulted;

stateLogic(ADR(_fireCount));
publishHMI();
flowLogic := TRUE;
END_METHOD

// AND-divergence: source done -> BOTH targets activate (parallel branches).
METHOD PROTECTED flowSplit2 : INT
VAR_INPUT
    inpFrom : INT;
    inpTo1  : INT;
    inpTo2  : INT;
    inpName : STRING(63) := '';
END_VAR
flowSplit2 := flow(inpFrom := inpFrom, inpTo := inpTo1, inpName := inpName);
IF flowSplit2 = 0 THEN
    RETURN;
END_IF
arcTo(inpTrans := flowSplit2, inpStepId := inpTo2);
END_METHOD

// AND-divergence: source done -> ALL THREE targets activate (parallel branches).
METHOD PROTECTED flowSplit3 : INT
VAR_INPUT
    inpFrom : INT;
    inpTo1  : INT;
    inpTo2  : INT;
    inpTo3  : INT;
    inpName : STRING(63) := '';
END_VAR
flowSplit3 := flow(inpFrom := inpFrom, inpTo := inpTo1, inpName := inpName);
IF flowSplit3 = 0 THEN
    RETURN;
END_IF
arcTo(inpTrans := flowSplit3, inpStepId := inpTo2);
arcTo(inpTrans := flowSplit3, inpStepId := inpTo3);
END_METHOD

METHOD PUBLIC getFlowHMIdata : ST_MachineFlow_HMI_Status
VAR_INPUT
END_VAR
getFlowHMIdata := HMIflow;
END_METHOD

METHOD PRIVATE placeToken : BOOL
VAR_INPUT
    inpStepId : INT;
END_VAR
_steps[inpStepId].active := TRUE;
_steps[inpStepId].done := FALSE;
_steps[inpStepId].entered := FALSE;
_steps[inpStepId].kickTimer := TRUE;   // restart the elapsed clock (also on re-entry)
placeToken := TRUE;
END_METHOD

METHOD PRIVATE publishHMI : BOOL
VAR_INPUT
END_VAR
VAR
    i     : INT;
    t     : INT;
    lo    : UDINT;
    hi    : UDINT;
    dLo   : UDINT;
    dHi   : UDINT;
    pLo   : UDINT;
    pHi   : UDINT;
    vLo   : UDINT;
    vHi   : UDINT;
    fLo   : UDINT;
    fHi   : UDINT;
    names : STRING(255);
    n     : INT;
END_VAR
FOR i := 1 TO _stepCount DO
    IF _steps[i].active THEN
        IF i <= 32 THEN
            lo := lo OR SHL(TO_UDINT(1), i - 1);
            IF _steps[i].done THEN
                dLo := dLo OR SHL(TO_UDINT(1), i - 1);
            END_IF
        ELSE
            hi := hi OR SHL(TO_UDINT(1), i - 33);
            IF _steps[i].done THEN
                dHi := dHi OR SHL(TO_UDINT(1), i - 33);
            END_IF
        END_IF
        IF n > 0 THEN
            names := CONCAT(names, ' + ');
        END_IF
        names := CONCAT(names, _steps[i].name);
        n := n + 1;
    END_IF
    // Outside the .active guard on purpose: a COMPLETED step has no token, so this bit is exactly
    // the information the active mask cannot carry.
    IF _steps[i].visited THEN
        IF i <= 32 THEN
            vLo := vLo OR SHL(TO_UDINT(1), i - 1);
        ELSE
            vHi := vHi OR SHL(TO_UDINT(1), i - 33);
        END_IF
    END_IF
END_FOR
FOR t := 1 TO _transCount DO
    // This mask IS the effective gate, because the boolean is: whatever ANDs into a transition's
    // permissive - a plain condition, an fb_Permissive's stsPermissiveOK, both - the machine ANDs in
    // before calling setPermissive(). Reporting a ready gate on a sequence that cannot advance would
    // be the exact symptom an operator is using the flow chart to diagnose.
    IF _trans[t].permissive THEN
        IF t <= 32 THEN
            pLo := pLo OR SHL(TO_UDINT(1), t - 1);
        ELSE
            pHi := pHi OR SHL(TO_UDINT(1), t - 33);
        END_IF
    END_IF
    IF _trans[t].fired THEN
        IF t <= 32 THEN
            fLo := fLo OR SHL(TO_UDINT(1), t - 1);
        ELSE
            fHi := fHi OR SHL(TO_UDINT(1), t - 33);
        END_IF
    END_IF
END_FOR
HMIflow.stsActiveLo := lo;
HMIflow.stsActiveHi := hi;
HMIflow.stsDoneLo := dLo;
HMIflow.stsDoneHi := dHi;
HMIflow.stsPermissiveLo := pLo;
HMIflow.stsPermissiveHi := pHi;
HMIflow.stsVisitedLo := vLo;
HMIflow.stsVisitedHi := vHi;
HMIflow.stsFiredLo := fLo;
HMIflow.stsFiredHi := fHi;
HMIflow.stsFaultedStep := _faultedStep;
HMIflow.stsFireCount := _fireCount;
HMIflow.stsLastFired := _lastFired;
stsActiveNames := names;
HMIflow.stsActiveNames := names;   // was declared but never written - see Docs/fb_MachineFlow_Design.md
IF stsRunning AND n > 0 THEN
    stsStepDescription := names;   // engine-owned while running
END_IF
publishHMI := TRUE;
END_METHOD

METHOD PRIVATE runStepTimers : BOOL
VAR_INPUT
END_VAR
VAR
    i : INT;
END_VAR
FOR i := 1 TO _stepCount DO
    // kickTimer forces one scan of IN=FALSE so the TON restarts on token placement
    _stepTimers[i](IN := _steps[i].active AND NOT _steps[i].kickTimer, PT := T#100H);
    IF _steps[i].kickTimer THEN
        _steps[i].kickTimer := FALSE;
    ELSIF _steps[i].active AND _steps[i].timeout > T#0S AND _stepTimers[i].ET > _steps[i].timeout THEN
        _timeoutStep := i;
        _faultedStep := i;   // a timeout is a step fault too — same red step on the chart
        setStateLogicFault(CONCAT('Step timeout: ', _steps[i].name), TRUE, _fireCount);
        RETURN;
    END_IF
END_FOR
runStepTimers := TRUE;
END_METHOD

METHOD PRIVATE seedTokens : BOOL
VAR_INPUT
END_VAR
VAR
    i : INT;
END_VAR
clearTokens();
_fireCount := 0;
_lastFired := 0;
_timeoutStep := 0;
_faultedStep := 0;
FOR i := 1 TO _stepCount DO
    IF _initialSteps[i] THEN
        placeToken(i);
    END_IF
END_FOR
seedTokens := TRUE;
END_METHOD

// Latch the FIRST definition error; actionsRun() faults on any run attempt.
// Report a CONFIGURATION error - a defineFlow() mistake, not a runtime fault. actionsRun turns it
// into a non-retryable fault, because a bad graph cannot be retried into a good one. PROTECTED so a
// subclass's defineFlow() can report its own (e.g. the addStep() id-drift guard in the header).
METHOD PROTECTED setCfgError : BOOL
VAR_INPUT
    inpMessage : STRING(255);
END_VAR
IF NOT _cfgError THEN
    _cfgError := TRUE;
    _cfgErrorText := inpMessage;
END_IF
setCfgError := TRUE;
END_METHOD

// Set a transition's permissive - the condition that must be MET to proceed
// (call from stepActions(), typically in the SOURCE step's body). Permissives
// are sticky and reset to TRUE on reset. OR-choice: opposing permissives on
// two transitions leaving the same step.
METHOD PROTECTED setPermissive : BOOL
VAR_INPUT
    inpTrans     : INT;
    inpCondition : BOOL;
END_VAR
IF inpTrans >= 1 AND inpTrans <= _transCount THEN
    _trans[inpTrans].permissive := inpCondition;
    setPermissive := TRUE;
END_IF
END_METHOD

// Mark a step as initially active on run (call from defineFlow(), AFTER the
// steps are declared; more than once for parallel starts). Default: step 1.
METHOD PROTECTED setInitialStep : BOOL
VAR_INPUT
    inpStepId : INT;
END_VAR
IF inpStepId < 1 OR inpStepId > _stepCount THEN
    setCfgError('MachineFlow: setInitialStep() unknown step');
    RETURN;
END_IF
IF NOT _initialSteps[inpStepId] THEN
    _initialSteps[inpStepId] := TRUE;
    _initialCount := _initialCount + 1;
END_IF
setInitialStep := TRUE;
END_METHOD

// Runtime timeout override (e.g. from a recipe) - replaces the addStep() value.
METHOD PROTECTED setStepTimeout : BOOL
VAR_INPUT
    inpStepId  : INT;
    inpTimeout : TIME;
END_VAR
IF inpStepId >= 1 AND inpStepId <= _stepCount THEN
    _steps[inpStepId].timeout := inpTimeout;
    setStepTimeout := TRUE;
END_IF
END_METHOD

// Override: the step BODIES - a CASE over the ids returned by addStep().
// Called once per ACTIVE step per scan (parallel steps each get their call);
// inpFirstScan is TRUE the first scan after the step's token arrives (use it
// for one-shot commands). Report completion with stepDone(inpStepId); fault
// via the inherited setStateLogicFault().
METHOD PROTECTED stepActions : BOOL
VAR_INPUT
    inpStepId    : INT;
    inpFirstScan : BOOL;
END_VAR
END_METHOD

METHOD PROTECTED stepActive : BOOL
VAR_INPUT
    inpStepId : INT;
END_VAR
IF inpStepId >= 1 AND inpStepId <= _stepCount THEN
    stepActive := _steps[inpStepId].active;
END_IF
END_METHOD

// Report a step complete (call from stepActions()). The token stays in place,
// marked done, until an outgoing transition consumes it - or, if the step has
// no outgoing transition, the sequence completes.
METHOD PROTECTED stepDone : BOOL
VAR_INPUT
    inpStepId : INT;
END_VAR
IF inpStepId >= 1 AND inpStepId <= _stepCount THEN
    IF _steps[inpStepId].active THEN
        _steps[inpStepId].done := TRUE;
        stepDone := TRUE;
    END_IF
END_IF
END_METHOD

// Time since this step's token arrived (each step has its own clock).
METHOD PROTECTED stepElapsed : TIME
VAR_INPUT
    inpStepId : INT;
END_VAR
IF inpStepId >= 1 AND inpStepId <= _stepCount THEN
    stepElapsed := _stepTimers[inpStepId].ET;
END_IF
END_METHOD

END_FUNCTION_BLOCK

// ---- POUs/FBs/Abstract/abs_fb_stateDevice.TcPOU
FUNCTION_BLOCK ABSTRACT abs_fb_stateDevice
VAR_INPUT
	inpReset	: BOOL;
	inpAuto		: BOOL;
	faultMonitor: POINTER TO fb_FaultMonitor;
END_VAR
VAR_OUTPUT
	stsIdle				: BOOL;
	stsDone				: BOOL;
	stsRunning			: BOOL;
	stsFaulted			: BOOL;
	stsAborting			: BOOL;
	stsAborted			: BOOL;
	stsFaultDescription	: STRING;
	stsStepDescription : STRING;
END_VAR
VAR
	_inAuto				: BOOL;
	_deviceName 		: STRING;
	_initMachineMode	: BOOL;
	_init				: BOOL;
	Interlock			: fb_Interlock;
	_dataInterlock		: st_interlock;
	// START permissive — the conditions that must be met to ENTER Running. Wire slots with
	// cmdSetStartPermissive(); unwired slots default TRUE, so an FB that never touches it is
	// satisfied and behaves exactly as before this was added.
	permStartPermissive	: fb_Permissive;
	_stateDoneAborting	: BOOL;
	_stateLogicReqRun	: BOOL;
	_stateLogicReset	: BOOL;
	_stateLogicFault	: FB_TcAlarm;
	_stateLogicMsg		: FB_TcMessage;
	_retryAllowed		: BOOL;
	_retryStep			: INT;
	_retryStateActive	: BOOL;
	_stateVariable		: POINTER TO INT;
	_lastStep			: INT;
	_stepTimer			: TON;
	_stepTimerEnable	: BOOL;
	_stepTimeoutPT		: TIME;
	HMIstateLogic		: ST_StateDevice_HMI_Interface;
	_stateLogicFaultRaised  : BOOL;
	_clear				: BOOL;
	_sentWarning		: STRING;
	_sentLog			: STRING;
	_runtimeTimer		: TON;
	_runtimeTimerTrig	: BOOL;
	_cycletime			: TIME;
	_cycletimeSet		: BOOL;
END_VAR

METHOD PROTECTED actionsAbort : BOOL
VAR_INPUT
END_VAR
END_METHOD

METHOD PROTECTED actionsDone : BOOL
VAR_INPUT
END_VAR
END_METHOD

METHOD PROTECTED actionsFaulted : BOOL
VAR_INPUT
END_VAR
END_METHOD

METHOD PROTECTED actionsReset : BOOL
VAR_INPUT
END_VAR
END_METHOD

METHOD PROTECTED actionsRun : BOOL
VAR_INPUT
END_VAR
END_METHOD

PROPERTY cfgDeviceName : STRING
GET
cfgDeviceName := _DeviceName;
END_GET
SET
_DeviceName := cfgDeviceName;
END_SET
END_PROPERTY

METHOD PUBLIC cmdSetInterlock : BOOL
VAR_INPUT
	interlockIndex : INT;
	description : STRING;
	condition: BOOL;
END_VAR
_dataInterlock.conditions[interlockIndex] := condition;
_dataInterlock.descriptions[interlockIndex] := description;
END_METHOD

// Wire one slot of the START permissive — a condition that must be met for this device to ENTER
// Running. Mirrors cmdSetInterlock's argument order on purpose, since a machine usually writes the
// two side by side; note fb_Permissive.setCondition() underneath takes (slot, met, description).
//
// Unwired slots default TRUE, so wire only what applies and leave the rest alone. Naming every slot
// you DO wire matters: that text is the operator's answer to "why won't it start".
//
// PERMISSIVE, NOT INTERLOCK: this gates the start only. A condition that must stop a device that is
// ALREADY RUNNING is an interlock — use cmdSetInterlock for that.
METHOD PUBLIC cmdSetStartPermissive : BOOL
VAR_INPUT
	inpSlot			: INT;
	inpDescription	: STRING;
	inpCondition	: BOOL;
END_VAR
cmdSetStartPermissive := permStartPermissive.setCondition(inpSlot, inpCondition, inpDescription);
END_METHOD

//FB_Init is always available implicitly and it is used primarily for initialization.
//The return value is not evaluated. For a specific influence, you can also declare the
//methods explicitly and provide additional code there with the standard initialization
//code. You can evaluate the return value.
METHOD FB_Init: BOOL
VAR_INPUT
    bInitRetains: BOOL; // TRUE: the retain variables are initialized (reset warm / reset cold)
    bInCopyCode: BOOL;  // TRUE: the instance will be copied to the copy code afterward (online change)
	cfgDeviceName 		: STRING;   
END_VAR
THIS^.cfgDeviceName 		:= 		cfgDeviceName;
END_METHOD

METHOD getStateLogicHMIdata : ST_StateDevice_HMI_Status
VAR_INPUT
END_VAR
getStateLogicHMIdata := HMIstateLogic.Status;
END_METHOD

METHOD sendLog : BOOL
VAR_INPUT
	message : STRING;
END_VAR
IF message <> _sentLog THEN
	_sentLog := message;
	_stateLogicMsg.CreateEx(TC_Events.absStateDevice.Logger,0);
	_stateLogicMsg.ipArguments.AddString(_deviceName).AddString(message);
	_stateLogicMsg.Send(0);
END_IF
END_METHOD

METHOD sendWarning : BOOL
VAR_INPUT
	message : STRING;
END_VAR
IF message <> _sentWarning THEN
	_sentWarning := message;
	_stateLogicMsg.CreateEx(TC_Events.absStateDevice.Warning,0);
	_stateLogicMsg.ipArguments.AddString(_deviceName).AddString(message);
	_stateLogicMsg.Send(0);	
END_IF
END_METHOD

METHOD INTERNAL setInit : BOOL
VAR_INPUT
END_VAR
IF faultMonitor <> 0 THEN
	faultMonitor^.addDeviceFault(faultStatus := ADR(stsFaulted), faultDescription := ADR(stsFaultDescription), deviceName := ADR(_deviceName));
END_IF
_stateLogicFault.CreateEx(stEventEntry:=TC_Events.absStateDevice.Faulted, bWithConfirmation := FALSE, ipSourceInfo := 0);
_stateLogicMsg.CreateEx(stEventEntry:=TC_events.absStateDevice.Warning,ipSourceInfo:=0);
_stateLogicMsg.CreateEx(stEventEntry:=TC_events.absStateDevice.Logger,ipSourceInfo:=0);
END_METHOD

METHOD setStateDoneAborting : BOOL
VAR_INPUT
END_VAR
_stateDoneAborting := TRUE;
END_METHOD

METHOD setStateLogicAbort : BOOL
VAR_INPUT
END_VAR
IF stsRunning THEN
	stsRunning := FALSE;
	stsAborting := TRUE;
END_IF
END_METHOD

METHOD setStateLogicDone : BOOL
VAR_INPUT
END_VAR
IF stsRunning THEN
	stsDone := TRUE;
END_IF
END_METHOD

METHOD setStateLogicFault : BOOL
VAR_INPUT
	FaultDescription : STRING;
	AllowRetry		 : BOOL;
	RetryStep		 : INT;
END_VAR
stsFaulted := TRUE;
stsFaultDescription := FaultDescription;

_retryAllowed := AllowRetry;
_retryStep	  := RetryStep;
END_METHOD

METHOD setStateLogicReset : BOOL
VAR_INPUT
END_VAR
_stateLogicReset := TRUE;
END_METHOD

METHOD setStateLogicRetry : BOOL
VAR_INPUT
END_VAR
IF stsFaulted THEN
	IF _retryAllowed THEN
		_retryStateActive := TRUE;
		_retryAllowed := FALSE;
		IF _stateVariable <> 0 THEN
			_stateVariable^ := _retryStep;
		END_IF
		stsFaulted := FALSE;
		stsFaultDescription := '';
		HMIstateLogic.Status.stsFaulted := FALSE;
		HMIstateLogic.Commands.ocmdRetry := FALSE;
		stsRunning := TRUE;
	END_IF
END_IF
END_METHOD

METHOD setStateLogicRun : BOOL
VAR_INPUT
END_VAR
IF stsIdle THEN
	_stateLogicReqRun := TRUE;
END_IF
END_METHOD

METHOD setStateLogicStepTimeout : BOOL
VAR_INPUT
	Timeout	: TIME;
END_VAR
IF _stepTimer.ET > Timeout THEN
	setStateLogicFault('Step timeout',TRUE,_stateVariable^);
	stsFaultDescription := concat('Step timeout on step ', INT_TO_STRING(_stateVariable^));
END_IF
END_METHOD

METHOD PROTECTED stateLogic : BOOL
VAR_INPUT
	stateVariable : POINTER TO INT;
END_VAR
IF NOT _init THEN
	_init := TRUE;
	setInit();
END_IF

_stateVariable := stateVariable;

//Measure duration of each step
_stepTimer(IN:= _stepTimerEnable, PT:= T#100H);

//Measure cycle time of the running state
_runtimeTimer(IN:=_runtimeTimerTrig, PT:=T#45D);
IF stsRunning THEN
	_runtimeTimerTrig := TRUE;
	_cycletimeset	  := FALSE;
	_cycletime:= _runtimeTimer.ET;
ELSE
	IF NOT(_cycletimeset) THEN
		_cycletimeset := TRUE;
		_cycletime:= _runtimeTimer.ET;
	END_IF
	_runtimetimerTrig := FALSE;	
END_IF

//Set interlocks
Interlock.name 			:= _DeviceName;
Interlock(inpConfig 	:= _dataInterlock);

// START permissive. Called HERE, before the run gate below, and unconditionally: stsPermissiveOK is
// a VAR_OUTPUT and reads FALSE until the body has run once, so gating on an uncalled instance would
// block every existing device on its first scan. Its conditions default TRUE, so an FB that never
// calls cmdSetStartPermissive() is satisfied from scan one.
permStartPermissive.cfgName := CONCAT(_DeviceName, ' start permissive');
permStartPermissive();

//Set Machine state
IF inpAuto THEN
	_inAuto := TRUE;
	HMIstateLogic.Status.stsAuto := TRUE;
ELSE
	_inAuto := FALSE;
	HMIstateLogic.Status.stsAuto := FALSE;
END_IF

//Run HMI operator commands if not in Auto
IF NOT(_inAuto) THEN
	IF HMIstateLogic.Commands.ocmdRun THEN
		setStateLogicRun();
	END_IF
	
	IF HMIstateLogic.Commands.ocmdAbort THEN
		setStateLogicAbort();
	END_IF
	
	IF HMIstateLogic.Commands.ocmdRetry THEN
		setStateLogicRetry();
	END_IF
	
END_IF

IF stsRunning OR stsFaulted OR stsDone OR stsAborted OR stsAborting THEN
	stsIdle 					 	:= FALSE;
	HMIstateLogic.Status.stsIdle 	:= FALSE;
ELSE
	stsIdle 						:= TRUE;
	HMIstateLogic.Status.stsIdle 	:= TRUE;
	HMIstateLogic.Status.stsState	:= 'Idle';
END_IF

IF HMIStateLogic.Commands.ocmdAbort THEN
	setStateLogicAbort();
END_IF

IF (inpReset OR HMIstatelogic.Commands.ocmdReset OR _stateLogicReset) AND (NOT(stsRunning) AND NOT(stsAborting)) THEN
	stsFaulted 								:= FALSE;
	stsAborted								:= FALSE;
	stsDone   								:= FALSE;
	stsRunning  							:= FALSE;
	stsIdle 								:= TRUE;
	HMIstateLogic.status.stsAborted			:= FALSE;
	HMIstateLogic.Status.stsFaulted 		:= FALSE;
	HMIstateLogic.Status.stsDone 			:= FALSE;
	HMIstateLogic.Status.stsRunning			:= FALSE;
	HMIstateLogic.Status.stsIdle 			:= TRUE;
	_stateLogicReset 						:= 0;
	_cycleTime								:= T#0s;
	stsStepDescription 	:= '';
	stsFaultDescription := '';

	IF _stateVariable <> 0 THEN
		_stateVariable^ 	:= 0;
	END_IF
	_retryStep				:= 0;
	_retryAllowed 			:= FALSE;
	
	IF NOT(stsFaulted) THEN
		_stateLogicFaultRaised := FALSE;
		_stateLogicFault.Clear(0);
	END_IF
	
	actionsReset();
ELSE
	_stateLogicReset := FALSE;
END_IF

IF stsAborting THEN
	HMIstateLogic.Status.stsRunning 		:= FALSE;
	_stateLogicReqRun						:= FALSE;
	stsStepDescription 						:= 'Aborting';
	HMIstateLogic.Status.stsState			:= 'Aborting';
	HMIstateLogic.Status.stsAborting		:= TRUE;
	IF _stateDoneAborting THEN
		stsAborting			 				:= FALSE;
		HMIstateLogic.Status.stsAborting	:= FALSE;
		stsAborted 			 				:= TRUE;
	END_IF
	actionsAbort();
END_IF

IF stsAborted THEN
	stsStepDescription 				:= 'Aborted';
	HMIstateLogic.Status.stsAborted := TRUE;
	HMIstateLogic.Status.stsState	:= 'Aborted';
	_stateDoneAborting				:= FALSE;
END_IF

IF stsFaulted THEN
	IF stsFaulted AND NOT(_stateLogicFaultRaised) THEN
		_stateLogicFaultRaised := TRUE;
		_stateLogicFault.ipArguments.Clear();
		_stateLogicFault.ipArguments.AddString(_deviceName).AddString(stsFaultDescription);
		_stateLogicFault.Raise(nTimeStamp :=0);
	END_IF
	stsRunning 			 			:= FALSE;
	HMIstateLogic.Status.stsRunning := FALSE;
	actionsFaulted();
	HMIstateLogic.Status.stsFaulted := TRUE;
	HMIstateLogic.Status.stsState	:= 'Faulted';
	_stepTimerEnable				:= FALSE;

END_IF

IF stsDone THEN
	_stateLogicReqRun 	:= FALSE;
	stsRunning := FALSE;
	actionsDone();
	HMIstateLogic.Status.stsRunning := FALSE;
	HMIstateLogic.Status.stsDone 	:= TRUE;
	HMIstateLogic.Status.stsState	:= 'Done';
END_IF

IF _stateLogicReqRun THEN
	IF stsIdle THEN
		IF NOT Interlock.outInterlockOK THEN
			sendWarning('Cannot start sequence, interlocks NOK');
		// A permissive gates the START and nothing else. It is deliberately NOT added to the
		// `IF stsRunning` check below, which aborts on a dropped INTERLOCK: an interlock breaking is
		// abnormal and must stop the device, whereas a permissive going unmet mid-run is normal and
		// means nothing — the device is already past the point it gated. Aborting on one would make
		// a permissive behave exactly like the interlock it exists to not be.
		ELSIF NOT permStartPermissive.stsPermissiveOK THEN
			sendWarning(CONCAT('Cannot start sequence, start permissive not met - unmet conditions: ',
				INT_TO_STRING(permStartPermissive.stsUnmetCount)));
		ELSE
			_stateLogicReqRun := FALSE;
			stsRunning := TRUE;
			_initMachineMode := _inAuto;
		END_IF
	ELSE
		sendWarning('Cannot start sequence, not in idle');
	END_IF
END_IF

IF stsRunning THEN
	IF NOT(Interlock.outInterlockOK) THEN
		sendWarning('Interlocks NOK, aborting...');
		setStateLogicAbort();
	ELSE
		_lastStep := _stateVariable^;
		_retryStateActive				:= FALSE;
		stsIdle 						:= FALSE;
		stsDone 						:= FALSE;
		stsRunning 						:= TRUE;
		HMIstateLogic.Status.stsRunning := TRUE;
		HMIstateLogic.Status.stsState	:= 'Running';
		actionsRun();
		//if Machine state changes from when running start (Auto to Man. or Man. to Auto) then abort
		IF _initMachineMode <> _inAuto THEN
			setStateLogicAbort();
		END_IF
		IF _stateVariable^ <> _lastStep THEN
			_stepTimerEnable := FALSE;
		ELSE
			_stepTimerEnable := TRUE;
		END_IF
	END_IF
ELSE
	_stateLogicReqRun := FALSE;
	_stepTimerEnable  := FALSE;
END_IF

HMIstateLogic.Status.cfgDeviceName 		 := _DeviceName;
HMIstateLogic.Status.stsStepDescription  := stsStepDescription;
HMIstateLogic.Status.stsFaultDescription := stsFaultDescription;
HMIstateLogic.Status.stsRetryAllowed	 := _retryAllowed;
HMIstateLogic.interlock 		  		 := Interlock.getHMIdata();
HMIstateLogic.startPermissive            := permStartPermissive.getHMIdata();
IF _stateVariable <> 0 THEN
	HMIstateLogic.Status.stsStepNumber := _stateVariable^;
END_IF

IF stsStepDescription <> '' THEN
	sendLog(stsStepDescription);
END_IF
END_METHOD

END_FUNCTION_BLOCK

// ---- POUs/FBs/fb_Permissive.TcPOU
(*
    fb_Permissive — a set of up to TEN conditions that must ALL be true for something to be
    ALLOWED to proceed. All-true means satisfied, and unwired slots default TRUE so you wire only
    what applies.

    SELF-CONTAINED, per CONVENTIONS §5: ten is a literal here, in ST_Permissive's array bounds and
    in the loops below — this FB references no GVL and reads no global state. Everything it needs
    arrives through inpConfig. Raising the capacity means editing those together.

    PERMISSIVE vs INTERLOCK — the distinction that decides which one you want:
      * an INTERLOCK (fb_Interlock) is a condition that must hold for a device to KEEP RUNNING.
        Breaking one is abnormal: it stops the device and it is a FAULT the operator must clear.
      * a PERMISSIVE is a condition that must be met for something to START or ADVANCE. Not being
        met yet is NORMAL — the machine is waiting, not broken. "Chamber not yet at vacuum" is not
        a fault, it is a Tuesday.
    So this FB deliberately raises NO fault, has no TcAlarm plumbing and does not extend
    abs_fb_Device. It answers exactly one question — "may this proceed, and if not, which conditions
    are not met".

    USAGE
        VAR
            PermStart : fb_Permissive;
        END_VAR

        // describe the slots once (startup or FB_Init of the owner)
        PermStart.inpConfig.descriptions[1] := 'Chamber door closed';
        PermStart.inpConfig.descriptions[2] := 'Vacuum below 5 Torr';
        PermStart.cfgName := 'Start permissive';

        // drive them every scan; leave unused slots alone (they stay TRUE)
        PermStart.inpConfig.conditions[1] := DoorClosed;
        PermStart.inpConfig.conditions[2] := Pressure < 5.0;
        PermStart();

        IF PermStart.stsPermissiveOK THEN ... END_IF

    NO FIRST-OUT, and that is the sharpest line between this and fb_Interlock. An interlock TRIPS:
    one condition drops, the device faults instantly, and "which one went first" names the cause -
    the later ones are usually consequences. A permissive never trips. It is simply evaluated at the
    moment something asks to proceed, and every unmet condition is equally and simultaneously the
    reason. There is no first, so the FB publishes the SET (stsConditions + stsUnmetCount) and the
    HMI shows all of them rather than nominating a misleading headline.

    NO BYPASS, either. It is tempting to allow one on the grounds that a permissive was never a
    safety function — but a bypass is precisely the control that makes an unsatisfied gate report
    itself satisfied, and a sequence advanced on a forced permissive fails later, somewhere that
    explains nothing. The conditions hold or they do not. If a condition needs to not apply, do not
    wire that slot; it defaults TRUE. (fb_Interlock's inpGlobalBypass is a genuinely different
    case: an interlock STOPS a running machine, so commissioning needs a documented way past it.)

    It is a DISPLAY-and-SEQUENCING aid, not a safety function: real safety lives in the safety PLC /
    hard wiring, and an interlock that must stop a running device belongs in fb_Interlock.

    Consumers: abs_fb_MachineFlow transition gates — the machine ANDs stsPermissiveOK into
    setPermissive(t, ...); MachineFlow holds no reference to this FB. Also device start conditions and
    the shared lhmi PermissiveList component (binds .HMI directly).
*)
FUNCTION_BLOCK fb_Permissive
VAR_INPUT
    inpConfig   : ST_Permissive;
END_VAR

VAR_OUTPUT
    stsPermissiveOK : BOOL;     // TRUE when every condition is met
    stsUnmetCount   : INT;      // number of unmet conditions
END_VAR

VAR
    i   : INT;
    HMI : ST_Permissive_HMI_Interface;
END_VAR

// Count every unmet slot every scan. The count is wanted even while satisfied, so there is no
// early exit.
//
// NO FIRST-OUT HERE, deliberately - see the header block. First-out is a TEMPORAL question and a
// permissive has no temporal dimension: nothing tripped, so no condition "went first". Every unmet
// condition is equally and simultaneously the reason, which is why the consumer shows the SET.
//
// 10 is a literal, matching ST_Permissive's array bound - CONVENTIONS §5. fb_Interlock's bound and
// its loop can drift apart for exactly this reason; keep these two edits together.
stsUnmetCount := 0;

FOR i := 1 TO 10 DO
    IF NOT inpConfig.conditions[i] THEN
        stsUnmetCount := stsUnmetCount + 1;
    END_IF
END_FOR

stsPermissiveOK := (stsUnmetCount = 0);

// ── publish to HMI (last section, per CONVENTIONS §3) ──
HMI.stsPermissiveOK := stsPermissiveOK;
HMI.stsConditions   := inpConfig.conditions;
HMI.stsDescriptions := inpConfig.descriptions;
HMI.stsUnmetCount   := stsUnmetCount;

METHOD PUBLIC getHMIdata : ST_Permissive_HMI_Interface
VAR_INPUT
END_VAR
getHMIdata := HMI;
END_METHOD

// Drive one slot, optionally naming it at the same time. Convenience over poking inpConfig
// directly: it bounds-checks the slot, so a typo'd index is a no-op instead of a memory scribble,
// and it keeps a condition and its description together at the call site where they are easiest to
// keep in step. Pass an empty inpDescription to leave the existing text alone.
METHOD PUBLIC setCondition : BOOL
VAR_INPUT
    inpSlot         : INT;
    inpMet          : BOOL;
    inpDescription  : STRING;
END_VAR
IF inpSlot < 1 OR inpSlot > 10 THEN
    setCondition := FALSE;
    RETURN;
END_IF

inpConfig.conditions[inpSlot] := inpMet;
IF inpDescription <> '' THEN
    inpConfig.descriptions[inpSlot] := inpDescription;
END_IF
setCondition := TRUE;
END_METHOD

// Operator-facing name for this permissive set, shown as the heading in the HMI list.
PROPERTY PUBLIC cfgName : STRING
GET
cfgName := HMI.stsPermissiveName;
END_GET
SET
HMI.stsPermissiveName := cfgName;
END_SET
END_PROPERTY

END_FUNCTION_BLOCK

// ---- POUs/FBs/Comm/fb_Modbus_Driver.TcPOU
// High-level Modbus TCP driver. Configuration-driven: define signals as
// arrays of ST_MBSignalConfig and the driver handles block optimization,
// endian conversion, RMW for bit-in-register writes, reconnection, and
// quality tracking.
//
// Usage:
//   1. Set properties (ipAddress, readSignalCount, writeSignalCount, ...)
//      BEFORE first enabling the FB.
//   2. Pass pointers to user arrays (config, results, write data) via inputs.
//   3. Call cycle() every PLC scan after the FB body call.
//   4. Optional: hold inpHoldWrites TRUE to keep reading without writing — e.g. until
//      the caller has read the device's current values to seed its write data from.
//
// Failure handling: after maxConsecFails failed transactions in a row the driver drops the
// link, waits reconnectDelay and retries; after maxReconnectAttempts such retries without a
// clean read cycle it stops in Faulted (no traffic) until cmdReset() or an enable toggle.
//
// Required library: Tc3_ModbusTCP (TF6250).
FUNCTION_BLOCK fb_Modbus_Driver
VAR_INPUT
    inpEnable               : BOOL;
    inpHoldWrites           : BOOL;     // TRUE = keep polling reads, start no write cycle

    inpPtrReadConfig        : POINTER TO ST_MBSignalConfig;
    inpPtrWriteConfig       : POINTER TO ST_MBSignalConfig;
    inpPtrReadResults       : POINTER TO ST_MBReadResult;
    inpPtrWriteData         : POINTER TO ST_MBWriteData;
END_VAR

VAR_OUTPUT
    stsStatus               : ST_MBDeviceStatus;
    stsError                : BOOL;
    stsErrorId              : UDINT;
END_VAR

VAR CONSTANT
    MAX_READ_SIGNALS        : UINT := 100;
    MAX_WRITE_SIGNALS       : UINT := 100;
    MAX_READ_BLOCKS         : UINT := 25;
    MAX_WRITE_BLOCKS        : UINT := 25;
    MAX_REGS_PER_BLOCK      : UINT := 125;
    MAX_COILS_PER_BLOCK     : UINT := 2000;
    MAX_SIGNALS_PER_BLOCK   : UINT := 64;
    MAX_BIT_REGISTERS       : UINT := 20;
    GAP_TOLERANCE_REGS      : UINT := 4;
    GAP_TOLERANCE_COILS     : UINT := 16;
    BIT_INDEX_NA            : BYTE := 255;
END_VAR

VAR
    // Configuration (set via properties before enable)
    cfgIpAddress            : STRING(15) := '192.168.1.1';
    cfgPort                 : UINT := 502;
    cfgUnitId               : BYTE := 1;
    cfgTimeout              : TIME := T#1S;
    cfgPollInterval         : TIME := T#100MS;
    cfgCommandDelay         : TIME := T#10MS;
    cfgWriteCycleInterval   : TIME := T#500MS;
    cfgWordOrder            : E_WordOrder := E_WordOrder.BigEndian;
    cfgMaxConsecFails       : UINT := 3;
    cfgStaleThreshold       : TIME := T#5S;
    cfgReconnectDelay       : TIME := T#2S;
    cfgMaxReconnectAttempts : UINT := 3;
    cfgReadSignalCount      : UINT;
    cfgWriteSignalCount     : UINT;

    // State machine
    _state                  : E_DriverState := E_DriverState.Init;
    _initialized            : BOOL;
    _enablePrev             : BOOL;

    // Connection state (Tc2_ModbusCaller manages TCP internally per FB call;
    // _socketConnected here means "driver is ready and last operation didn't fail")
    _socketConnected        : BOOL;
    _connectAttempts        : UINT;
    _disconnectPending      : BOOL;

    // Timing
    tonPollInterval         : TON;
    tonWriteInterval        : TON;
    tonCommandDelay         : TON;
    tonTimeout              : TON;
    tonReconnectDelay       : TON;
    _lastGoodReadTime       : TIME;
    _lastGoodWriteTime      : TIME;

    // Parsed configuration
    _arrParsedRead          : ARRAY[1..100] OF ST_ParsedSignal;
    _arrParsedWrite         : ARRAY[1..100] OF ST_ParsedSignal;

    // Optimized blocks
    _arrReadBlocks          : ARRAY[1..25] OF ST_ReadBlock;
    _readBlockCount         : UINT;

    _arrWriteBlocks         : ARRAY[1..25] OF ST_WriteBlock;
    _writeBlockCount        : UINT;

    // Bit register tracking (RMW)
    _arrBitRegisters        : ARRAY[1..20] OF ST_BitRegisterRmw;
    _bitRegisterCount       : UINT;

    // Runtime indices
    _currentBlockIdx        : UINT;
    _currentRmwIdx          : UINT;

    // Raw data buffers
    _arrRawReadBuffer       : ARRAY[0..124] OF WORD;
    _arrRawWriteBuffer      : ARRAY[0..124] OF WORD;

    // Tc2_ModbusCaller function blocks (each manages its own TCP connection)
    fbMbReadCoils           : FB_MBReadCoils;       // FC01
    fbMbReadInputs          : FB_MBReadInputs;      // FC02 (discrete inputs)
    fbMbReadRegs            : FB_MBReadRegs;        // FC03 (holding regs)
    fbMbReadInputRegs       : FB_MBReadInputRegs;   // FC04 (input regs)
    fbMbWriteSingleCoil     : FB_MBWriteSingleCoil; // FC05
    fbMbWriteSingleReg      : FB_MBWriteSingleReg;  // FC06
    fbMbWriteCoils          : FB_MBWriteCoils;      // FC15
    fbMbWriteRegs           : FB_MBWriteRegs;       // FC16

    // Error tracking
    _consecFailures         : UINT;
    _lastMbError            : UDINT;
    _readCycleFailed        : BOOL;     // a block failed in the current read cycle
    _writeCycleFailed       : BOOL;     // a block failed in the current write cycle
    _resetRequest           : BOOL;     // cmdReset(): restart from Init without an enable edge

    // Sorting workspace
    _arrSortIdx             : ARRAY[1..100] OF UINT;
END_VAR

// FB body intentionally empty. All work is performed in the cycle() method,
// which the user must call once per PLC scan after invoking the FB itself.
;

METHOD PRIVATE applyBitModifications
VAR_INPUT
    inpRmwIdx : UINT;
END_VAR
VAR
    _reg        : REFERENCE TO ST_BitRegisterRmw;
    _baseValue  : WORD;
    _bitIdx     : UINT;
    _sigIdx     : UINT;
    _pData      : POINTER TO ST_MBWriteData;
END_VAR
_reg REF= _arrBitRegisters[inpRmwIdx];

_baseValue := swapBytes(_reg.readValue);

